// TIA Portal project "PLC_SWaT_LSTM" (V19)
// zoltan.dobrady@hotmail.com

(* hardware
DEVICE "S7-1500/ET200MP station_1"  S7-1500 station
   slot 0: "Rail_0"  Rack  6ES7 590-1***0-0AA0
   slot 1: "PLC_1"  CPU 1515F-2 PN  6ES7 515-2FM01-0AB0  V2.1
      slot 3: "CPU display_1"  6ES7591-1BA00-0AA0
      slot 32768: "PROFINET interface_1"  X1
         slot 32769: "Port_1"  X1 P1
         slot 32770: "Port_2"  X1 P2
      slot 33024: "PROFINET interface_2"  X2
         slot 33025: "Port_1"  X2 P1
*)

// ===== PLC "PLC_1"  CPU 1515F-2 PN =====

// folder: Database

DATA_BLOCK "DB_model_HS16_IW10"   // DB1
{ S7_Optimized_Access := 'TRUE' }
VERSION : 0.1
// --- Siemens Structured Format ---
   VAR
      W_i : Array[0..15, 0..39] of Real;
      W_f : Array[0..15, 0..39] of Real;
      W_g : Array[0..15, 0..39] of Real;
      W_o : Array[0..15, 0..39] of Real;
      R_i : Array[0..15, 0..15] of Real;
      R_f : Array[0..15, 0..15] of Real;
      R_g : Array[0..15, 0..15] of Real;
      R_o : Array[0..15, 0..15] of Real;
      B_i : Array[0..15] of Real;
      B_f : Array[0..15] of Real;
      B_g : Array[0..15] of Real;
      B_o : Array[0..15] of Real;
      FC_W : Array[0..39, 0..15] of Real;
      FC_B : Array[0..39] of Real;
   END_VAR
BEGIN
   W_i[0,0] := 0.03254747;
   W_i[0,1] := 0.123859;
   W_i[0,2] := 0.04015401;
   W_i[0,3] := -0.03803189;
   W_i[0,4] := 0.1759319;
   W_i[0,5] := 0.00417833;
   W_i[0,6] := -0.00157293;
   W_i[0,7] := 0.0728622;
   W_i[0,8] := 0.06175515;
   W_i[0,9] := -0.03080547;
   W_i[0,10] := 0.01361996;
   W_i[0,11] := -0.2367004;
   W_i[0,12] := 0.1251248;
   W_i[0,13] := -0.1203895;
   W_i[0,14] := 0.0523482;
   W_i[0,15] := 0.2630532;
   W_i[0,16] := -0.1147504;
   W_i[0,17] := 0.05957858;
   W_i[0,18] := -0.02271187;
   W_i[0,19] := -0.04982074;
   W_i[0,20] := 0.01270425;
   W_i[0,21] := 0.3620531;
   W_i[0,22] := -0.2914467;
   W_i[0,23] := 0.02366253;
   W_i[0,24] := -0.602429;
   W_i[0,25] := -0.5198534;
   W_i[0,26] := 0.01890776;
   W_i[0,27] := -0.4244256;
   W_i[0,28] := 0.09802054;
   W_i[0,29] := -0.2919731;
   W_i[0,30] := 0.1756448;
   W_i[0,31] := -0.06584074;
   W_i[0,32] := 0.04272554;
   W_i[0,33] := 0.06813997;
   W_i[0,34] := 0.1243908;
   W_i[0,35] := -0.2062567;
   W_i[0,36] := 0.05875245;
   W_i[0,37] := -0.2700093;
   W_i[0,38] := 0.2212317;
   W_i[0,39] := 1.454268;
   W_i[1,0] := 0.04402059;
   W_i[1,1] := 0.1007617;
   W_i[1,2] := -0.00997876;
   W_i[1,3] := 0.00796912;
   W_i[1,4] := -0.00383734;
   W_i[1,5] := -0.00800767;
   W_i[1,6] := 0.1229124;
   W_i[1,7] := 0.04417216;
   W_i[1,8] := -0.00160155;
   W_i[1,9] := -0.03973384;
   W_i[1,10] := -0.05576275;
   W_i[1,11] := 0.01415846;
   W_i[1,12] := -0.1102211;
   W_i[1,13] := 0.0361371;
   W_i[1,14] := -0.00464776;
   W_i[1,15] := -0.02071899;
   W_i[1,16] := 0.0165178;
   W_i[1,17] := -0.00011115;
   W_i[1,18] := 0.04986879;
   W_i[1,19] := -0.05042609;
   W_i[1,20] := 0.08610544;
   W_i[1,21] := 0.05673008;
   W_i[1,22] := -0.00434864;
   W_i[1,23] := 0.01197722;
   W_i[1,24] := -0.5458539;
   W_i[1,25] := -0.6899631;
   W_i[1,26] := 0.01104975;
   W_i[1,27] := 0.0182511;
   W_i[1,28] := 0.04478757;
   W_i[1,29] := -0.05586376;
   W_i[1,30] := 0.02979602;
   W_i[1,31] := 0.00707946;
   W_i[1,32] := 0.1464935;
   W_i[1,33] := 0.04832766;
   W_i[1,34] := -0.9202742;
   W_i[1,35] := -0.1918912;
   W_i[1,36] := 0.02485085;
   W_i[1,37] := -0.05241579;
   W_i[1,38] := 0.01553158;
   W_i[1,39] := -0.00394726;
   W_i[2,0] := 0.0670436;
   W_i[2,1] := -0.1175203;
   W_i[2,2] := 0.02326228;
   W_i[2,3] := -0.1431773;
   W_i[2,4] := -0.05582308;
   W_i[2,5] := 0.03605313;
   W_i[2,6] := 0.04952687;
   W_i[2,7] := -0.05419854;
   W_i[2,8] := -0.00077774;
   W_i[2,9] := 0.1769989;
   W_i[2,10] := 0.02469403;
   W_i[2,11] := 0.2849406;
   W_i[2,12] := -0.2712711;
   W_i[2,13] := -0.06837726;
   W_i[2,14] := 0.00509281;
   W_i[2,15] := 0.07467768;
   W_i[2,16] := 0.01470727;
   W_i[2,17] := 0.1139419;
   W_i[2,18] := -0.03895494;
   W_i[2,19] := 0.02999579;
   W_i[2,20] := 0.0196714;
   W_i[2,21] := 0.00220801;
   W_i[2,22] := -0.33803;
   W_i[2,23] := 0.09799825;
   W_i[2,24] := -0.5955718;
   W_i[2,25] := -0.7228485;
   W_i[2,26] := 0.07928592;
   W_i[2,27] := -0.03053538;
   W_i[2,28] := -0.1309938;
   W_i[2,29] := -0.04490006;
   W_i[2,30] := 0.05262627;
   W_i[2,31] := -0.03356259;
   W_i[2,32] := 0.06378829;
   W_i[2,33] := -0.00362085;
   W_i[2,34] := -0.6579466;
   W_i[2,35] := 0.02030313;
   W_i[2,36] := 0.05807094;
   W_i[2,37] := -0.1117615;
   W_i[2,38] := 0.09806133;
   W_i[2,39] := -0.04513157;
   W_i[3,0] := -0.03288125;
   W_i[3,1] := 0.03644303;
   W_i[3,2] := -0.02111984;
   W_i[3,3] := -0.09554495;
   W_i[3,4] := 0.471034;
   W_i[3,5] := -0.0182176;
   W_i[3,6] := -0.01296977;
   W_i[3,7] := 0.09772011;
   W_i[3,8] := 0.02375359;
   W_i[3,9] := 0.0802948;
   W_i[3,10] := 0.06341432;
   W_i[3,11] := -0.05777879;
   W_i[3,12] := 0.09200994;
   W_i[3,13] := -0.0054342;
   W_i[3,14] := -0.1107964;
   W_i[3,15] := 0.1856784;
   W_i[3,16] := -0.0179559;
   W_i[3,17] := -0.01424691;
   W_i[3,18] := 0.02418556;
   W_i[3,19] := -0.08783326;
   W_i[3,20] := 0.05560731;
   W_i[3,21] := 0.2986822;
   W_i[3,22] := -0.2220259;
   W_i[3,23] := -0.03734203;
   W_i[3,24] := 0.08825689;
   W_i[3,25] := 0.1838893;
   W_i[3,26] := 0.1152585;
   W_i[3,27] := -0.444976;
   W_i[3,28] := 0.1019801;
   W_i[3,29] := -0.4402614;
   W_i[3,30] := -0.2070405;
   W_i[3,31] := 0.00454621;
   W_i[3,32] := -0.03864358;
   W_i[3,33] := -0.1032195;
   W_i[3,34] := 0.6178231;
   W_i[3,35] := -0.01621445;
   W_i[3,36] := 0.06078746;
   W_i[3,37] := 0.07829241;
   W_i[3,38] := 0.08872399;
   W_i[3,39] := 0.01815886;
   W_i[4,0] := -0.09336383;
   W_i[4,1] := 0.00870158;
   W_i[4,2] := -0.0504511;
   W_i[4,3] := 0.0685437;
   W_i[4,4] := 0.06657482;
   W_i[4,5] := -0.04358229;
   W_i[4,6] := 0.01173393;
   W_i[4,7] := 0.02832152;
   W_i[4,8] := -0.2380867;
   W_i[4,9] := 0.2590344;
   W_i[4,10] := -0.02959821;
   W_i[4,11] := -0.1970284;
   W_i[4,12] := -0.04782372;
   W_i[4,13] := 0.00693473;
   W_i[4,14] := 0.00193878;
   W_i[4,15] := 0.03396931;
   W_i[4,16] := -0.03933699;
   W_i[4,17] := -0.09345319;
   W_i[4,18] := 0.8571873;
   W_i[4,19] := -0.208394;
   W_i[4,20] := -0.00447866;
   W_i[4,21] := -0.04350503;
   W_i[4,22] := 0.09176219;
   W_i[4,23] := 0.04992297;
   W_i[4,24] := -0.4504299;
   W_i[4,25] := 0.01641427;
   W_i[4,26] := -0.1837832;
   W_i[4,27] := 0.03955682;
   W_i[4,28] := -0.06913128;
   W_i[4,29] := 0.08025265;
   W_i[4,30] := -0.1162292;
   W_i[4,31] := 0.04558431;
   W_i[4,32] := 0.07176397;
   W_i[4,33] := -0.04032118;
   W_i[4,34] := 0.2098121;
   W_i[4,35] := -0.1125335;
   W_i[4,36] := -0.01868857;
   W_i[4,37] := -0.07242457;
   W_i[4,38] := -0.1324239;
   W_i[4,39] := -0.04244877;
   W_i[5,0] := 0.01391891;
   W_i[5,1] := -0.110183;
   W_i[5,2] := -0.00893384;
   W_i[5,3] := -0.01407803;
   W_i[5,4] := 0.08575681;
   W_i[5,5] := 0.08241521;
   W_i[5,6] := -0.06153676;
   W_i[5,7] := 0.03060099;
   W_i[5,8] := -0.03490681;
   W_i[5,9] := 0.0314279;
   W_i[5,10] := -0.02459875;
   W_i[5,11] := 0.1095907;
   W_i[5,12] := -0.02965787;
   W_i[5,13] := 0.00184801;
   W_i[5,14] := 0.02055808;
   W_i[5,15] := -0.00937524;
   W_i[5,16] := -0.01257727;
   W_i[5,17] := 0.01791891;
   W_i[5,18] := -0.0115625;
   W_i[5,19] := -0.02731706;
   W_i[5,20] := 0.08900256;
   W_i[5,21] := 0.09895428;
   W_i[5,22] := 0.02720478;
   W_i[5,23] := 0.04369688;
   W_i[5,24] := -1.906074;
   W_i[5,25] := -0.09418426;
   W_i[5,26] := -0.010597;
   W_i[5,27] := -0.09780212;
   W_i[5,28] := 0.1125583;
   W_i[5,29] := 0.08197493;
   W_i[5,30] := -0.08072126;
   W_i[5,31] := 0.03083795;
   W_i[5,32] := 0.06895962;
   W_i[5,33] := 0.00149198;
   W_i[5,34] := 0.3009818;
   W_i[5,35] := 0.1442458;
   W_i[5,36] := -0.02817895;
   W_i[5,37] := -0.08498497;
   W_i[5,38] := 0.03758771;
   W_i[5,39] := 0.01095005;
   W_i[6,0] := 0.08324189;
   W_i[6,1] := -0.2883669;
   W_i[6,2] := -0.00092833;
   W_i[6,3] := -0.00874277;
   W_i[6,4] := 0.1196982;
   W_i[6,5] := -0.1120785;
   W_i[6,6] := -0.0087709;
   W_i[6,7] := -0.03745995;
   W_i[6,8] := 0.00287988;
   W_i[6,9] := 0.00178848;
   W_i[6,10] := 0.03823818;
   W_i[6,11] := 0.02621512;
   W_i[6,12] := -0.288421;
   W_i[6,13] := -0.07084718;
   W_i[6,14] := 0.04070705;
   W_i[6,15] := -0.020424;
   W_i[6,16] := -0.00164282;
   W_i[6,17] := 0.01065832;
   W_i[6,18] := 0.00655926;
   W_i[6,19] := 0.02358968;
   W_i[6,20] := 0.1303789;
   W_i[6,21] := 0.038681;
   W_i[6,22] := -0.06235948;
   W_i[6,23] := 0.07983913;
   W_i[6,24] := -0.2428008;
   W_i[6,25] := -0.05732525;
   W_i[6,26] := 0.1651715;
   W_i[6,27] := -0.07414961;
   W_i[6,28] := 0.06032364;
   W_i[6,29] := 0.08282514;
   W_i[6,30] := -0.01358633;
   W_i[6,31] := 0.0431109;
   W_i[6,32] := 0.03472897;
   W_i[6,33] := -0.04253995;
   W_i[6,34] := 0.01447233;
   W_i[6,35] := 0.03594886;
   W_i[6,36] := -0.01385077;
   W_i[6,37] := 0.1116451;
   W_i[6,38] := 0.1253235;
   W_i[6,39] := -0.03726343;
   W_i[7,0] := 0.01927893;
   W_i[7,1] := 0.05625859;
   W_i[7,2] := 0.04672581;
   W_i[7,3] := -0.00316564;
   W_i[7,4] := 0.09401099;
   W_i[7,5] := -0.02755413;
   W_i[7,6] := -0.03952036;
   W_i[7,7] := 0.03364034;
   W_i[7,8] := 0.05500693;
   W_i[7,9] := 0.02471298;
   W_i[7,10] := 0.03820876;
   W_i[7,11] := -0.2692161;
   W_i[7,12] := -0.02231521;
   W_i[7,13] := -0.0175243;
   W_i[7,14] := 0.03934914;
   W_i[7,15] := 0.01282423;
   W_i[7,16] := -0.0871601;
   W_i[7,17] := -0.09125534;
   W_i[7,18] := 0.00613662;
   W_i[7,19] := 0.08651425;
   W_i[7,20] := -0.01288831;
   W_i[7,21] := 0.2017677;
   W_i[7,22] := -0.2016672;
   W_i[7,23] := 0.01241351;
   W_i[7,24] := -0.8755623;
   W_i[7,25] := -0.4621839;
   W_i[7,26] := 0.09773878;
   W_i[7,27] := -0.1281056;
   W_i[7,28] := 0.04194518;
   W_i[7,29] := -0.03563948;
   W_i[7,30] := 0.08049577;
   W_i[7,31] := 0.04509509;
   W_i[7,32] := -0.113328;
   W_i[7,33] := 0.1053996;
   W_i[7,34] := 0.2416716;
   W_i[7,35] := 0.04508473;
   W_i[7,36] := 0.00324964;
   W_i[7,37] := 0.2255004;
   W_i[7,38] := 0.1750992;
   W_i[7,39] := -0.7787634;
   W_i[8,0] := -0.03076644;
   W_i[8,1] := 0.03958185;
   W_i[8,2] := 0.05958826;
   W_i[8,3] := 0.00143461;
   W_i[8,4] := -0.03551066;
   W_i[8,5] := 0.0670559;
   W_i[8,6] := -0.00545013;
   W_i[8,7] := -0.1152002;
   W_i[8,8] := -0.04941865;
   W_i[8,9] := 0.00970779;
   W_i[8,10] := -0.02700928;
   W_i[8,11] := 0.1261697;
   W_i[8,12] := -0.230127;
   W_i[8,13] := -0.1321811;
   W_i[8,14] := 0.1056539;
   W_i[8,15] := 0.03265957;
   W_i[8,16] := 0.01893855;
   W_i[8,17] := 0.05783269;
   W_i[8,18] := 0.04541522;
   W_i[8,19] := -0.1756509;
   W_i[8,20] := -0.0300831;
   W_i[8,21] := 0.02609591;
   W_i[8,22] := -0.1179207;
   W_i[8,23] := -0.03097328;
   W_i[8,24] := -1.123494;
   W_i[8,25] := -0.1057856;
   W_i[8,26] := 0.1196709;
   W_i[8,27] := -0.1930985;
   W_i[8,28] := -0.04314341;
   W_i[8,29] := -0.02280886;
   W_i[8,30] := 0.09419166;
   W_i[8,31] := -0.00168002;
   W_i[8,32] := 0.170113;
   W_i[8,33] := 0.1277638;
   W_i[8,34] := 0.0079219;
   W_i[8,35] := 0.00793266;
   W_i[8,36] := 0.02933485;
   W_i[8,37] := -0.04765635;
   W_i[8,38] := -0.05385318;
   W_i[8,39] := 1.045761;
   W_i[9,0] := 0.1591891;
   W_i[9,1] := 0.04106269;
   W_i[9,2] := 0.02940365;
   W_i[9,3] := -0.02633034;
   W_i[9,4] := 0.06646424;
   W_i[9,5] := -0.06870057;
   W_i[9,6] := 0.00617184;
   W_i[9,7] := 0.01493581;
   W_i[9,8] := 0.00472299;
   W_i[9,9] := -0.1817109;
   W_i[9,10] := -0.0086358;
   W_i[9,11] := 0.1120397;
   W_i[9,12] := 0.03235663;
   W_i[9,13] := -0.00635904;
   W_i[9,14] := -0.00805719;
   W_i[9,15] := 0.03256573;
   W_i[9,16] := -0.029828;
   W_i[9,17] := 0.02432551;
   W_i[9,18] := -0.04791717;
   W_i[9,19] := -0.03479305;
   W_i[9,20] := 0.02419964;
   W_i[9,21] := -0.0080657;
   W_i[9,22] := 0.00884045;
   W_i[9,23] := 0.00822151;
   W_i[9,24] := -0.4626606;
   W_i[9,25] := -0.2415425;
   W_i[9,26] := 0.1063772;
   W_i[9,27] := 0.00555547;
   W_i[9,28] := 0.00231378;
   W_i[9,29] := 0.1730648;
   W_i[9,30] := -0.1442872;
   W_i[9,31] := -0.01611738;
   W_i[9,32] := -0.1527355;
   W_i[9,33] := -0.03995335;
   W_i[9,34] := -0.6023377;
   W_i[9,35] := -0.06071381;
   W_i[9,36] := 0.01153921;
   W_i[9,37] := 0.157252;
   W_i[9,38] := 0.04887648;
   W_i[9,39] := 0.03194974;
   W_i[10,0] := 5.71E-06;
   W_i[10,1] := 0.0292189;
   W_i[10,2] := 0.03921259;
   W_i[10,3] := -0.1034236;
   W_i[10,4] := 0.04451175;
   W_i[10,5] := -0.01788418;
   W_i[10,6] := 0.06014212;
   W_i[10,7] := -0.127616;
   W_i[10,8] := 0.1096968;
   W_i[10,9] := 0.1346427;
   W_i[10,10] := -0.07629871;
   W_i[10,11] := -1.314735;
   W_i[10,12] := 0.9704102;
   W_i[10,13] := -0.02917644;
   W_i[10,14] := 0.2685799;
   W_i[10,15] := 0.06801854;
   W_i[10,16] := -0.2241947;
   W_i[10,17] := 0.2624845;
   W_i[10,18] := -0.1694944;
   W_i[10,19] := -0.1197102;
   W_i[10,20] := -0.1591434;
   W_i[10,21] := 0.1818019;
   W_i[10,22] := -0.4487775;
   W_i[10,23] := 0.05718501;
   W_i[10,24] := 0.7740152;
   W_i[10,25] := 0.6112806;
   W_i[10,26] := 0.00735129;
   W_i[10,27] := -0.08243502;
   W_i[10,28] := -0.03729297;
   W_i[10,29] := 0.1612841;
   W_i[10,30] := -0.02351914;
   W_i[10,31] := 0.1043125;
   W_i[10,32] := 0.05746254;
   W_i[10,33] := 0.08887602;
   W_i[10,34] := -0.3910645;
   W_i[10,35] := 0.2256924;
   W_i[10,36] := -0.1320819;
   W_i[10,37] := -0.1611588;
   W_i[10,38] := 0.2708046;
   W_i[10,39] := 0.6280136;
   W_i[11,0] := -0.05849513;
   W_i[11,1] := -0.03062119;
   W_i[11,2] := -0.00411083;
   W_i[11,3] := 0.00799791;
   W_i[11,4] := 0.08333463;
   W_i[11,5] := 0.02937987;
   W_i[11,6] := 0.06844535;
   W_i[11,7] := -0.0119828;
   W_i[11,8] := 0.05660131;
   W_i[11,9] := -0.1460933;
   W_i[11,10] := -0.01666861;
   W_i[11,11] := -0.06908122;
   W_i[11,12] := 0.1548331;
   W_i[11,13] := -0.00687739;
   W_i[11,14] := 0.01971146;
   W_i[11,15] := 0.1330592;
   W_i[11,16] := -0.02189317;
   W_i[11,17] := 0.00985993;
   W_i[11,18] := -0.1488067;
   W_i[11,19] := 0.01909257;
   W_i[11,20] := 0.03714932;
   W_i[11,21] := -0.02673176;
   W_i[11,22] := -0.02788893;
   W_i[11,23] := 0.1140895;
   W_i[11,24] := -0.3711884;
   W_i[11,25] := -0.08985706;
   W_i[11,26] := -0.1102327;
   W_i[11,27] := 0.05117378;
   W_i[11,28] := 0.08547711;
   W_i[11,29] := 0.1270248;
   W_i[11,30] := 0.1054488;
   W_i[11,31] := -0.00480978;
   W_i[11,32] := 0.1614495;
   W_i[11,33] := 0.05210381;
   W_i[11,34] := -0.00085451;
   W_i[11,35] := -0.00874526;
   W_i[11,36] := -0.0616112;
   W_i[11,37] := -0.3677483;
   W_i[11,38] := 0.04212995;
   W_i[11,39] := 0.03037546;
   W_i[12,0] := 0.00629061;
   W_i[12,1] := -0.06136212;
   W_i[12,2] := -0.00718669;
   W_i[12,3] := -0.1004218;
   W_i[12,4] := 0.06293897;
   W_i[12,5] := -0.03143417;
   W_i[12,6] := -0.03538829;
   W_i[12,7] := 0.07763195;
   W_i[12,8] := -0.01023159;
   W_i[12,9] := -0.1141296;
   W_i[12,10] := -0.01354402;
   W_i[12,11] := -0.02311977;
   W_i[12,12] := 0.0279608;
   W_i[12,13] := 0.07165248;
   W_i[12,14] := -0.03632027;
   W_i[12,15] := 0.03878558;
   W_i[12,16] := -0.073125;
   W_i[12,17] := 0.01845204;
   W_i[12,18] := -0.08527449;
   W_i[12,19] := -0.00854577;
   W_i[12,20] := 0.00351815;
   W_i[12,21] := -0.1662848;
   W_i[12,22] := 0.06705266;
   W_i[12,23] := 0.1430702;
   W_i[12,24] := -0.539574;
   W_i[12,25] := -0.8721982;
   W_i[12,26] := -0.06440469;
   W_i[12,27] := 0.07379381;
   W_i[12,28] := 0.07828815;
   W_i[12,29] := 0.3882209;
   W_i[12,30] := 0.1159498;
   W_i[12,31] := 0.05581488;
   W_i[12,32] := 0.3066402;
   W_i[12,33] := 0.1275958;
   W_i[12,34] := -0.147978;
   W_i[12,35] := 0.1432935;
   W_i[12,36] := 0.2298153;
   W_i[12,37] := 0.00895516;
   W_i[12,38] := 0.2001298;
   W_i[12,39] := 0.09707437;
   W_i[13,0] := 0.07871004;
   W_i[13,1] := 0.0640982;
   W_i[13,2] := -0.00181766;
   W_i[13,3] := 0.05780525;
   W_i[13,4] := 0.2101672;
   W_i[13,5] := 0.05360549;
   W_i[13,6] := -0.0875827;
   W_i[13,7] := -0.3342811;
   W_i[13,8] := -0.09135646;
   W_i[13,9] := 0.1170631;
   W_i[13,10] := -0.0523126;
   W_i[13,11] := -0.03317479;
   W_i[13,12] := -0.403383;
   W_i[13,13] := -0.00985299;
   W_i[13,14] := 0.02202887;
   W_i[13,15] := 0.130378;
   W_i[13,16] := 0.04808246;
   W_i[13,17] := 0.04501719;
   W_i[13,18] := -0.01153503;
   W_i[13,19] := 0.03141625;
   W_i[13,20] := 0.02999944;
   W_i[13,21] := 0.01402024;
   W_i[13,22] := 0.06788336;
   W_i[13,23] := -0.09942459;
   W_i[13,24] := 0.3184399;
   W_i[13,25] := 0.1069793;
   W_i[13,26] := -0.06989229;
   W_i[13,27] := 0.1058815;
   W_i[13,28] := 0.06872193;
   W_i[13,29] := -0.1537144;
   W_i[13,30] := 0.06626805;
   W_i[13,31] := -0.0559484;
   W_i[13,32] := -0.09573574;
   W_i[13,33] := 0.05669653;
   W_i[13,34] := 0.06202357;
   W_i[13,35] := -0.1367418;
   W_i[13,36] := 0.06451428;
   W_i[13,37] := 0.1204168;
   W_i[13,38] := -0.168509;
   W_i[13,39] := 0.9775926;
   W_i[14,0] := 0.00773311;
   W_i[14,1] := -0.06673568;
   W_i[14,2] := -0.03463669;
   W_i[14,3] := -0.07830913;
   W_i[14,4] := 0.22799;
   W_i[14,5] := -0.2344869;
   W_i[14,6] := 0.1956936;
   W_i[14,7] := 0.1315334;
   W_i[14,8] := -0.1242086;
   W_i[14,9] := 0.2860397;
   W_i[14,10] := -0.09231006;
   W_i[14,11] := -0.2547791;
   W_i[14,12] := 0.1490363;
   W_i[14,13] := -0.2912802;
   W_i[14,14] := 0.1072571;
   W_i[14,15] := 0.1354038;
   W_i[14,16] := -0.09035023;
   W_i[14,17] := -0.01749873;
   W_i[14,18] := -0.4789497;
   W_i[14,19] := -0.06870104;
   W_i[14,20] := -0.1709639;
   W_i[14,21] := -0.05212005;
   W_i[14,22] := -0.1618474;
   W_i[14,23] := -0.2139406;
   W_i[14,24] := -0.7570689;
   W_i[14,25] := -0.7048593;
   W_i[14,26] := -0.3352102;
   W_i[14,27] := 0.03507431;
   W_i[14,28] := -0.1267896;
   W_i[14,29] := 0.1670964;
   W_i[14,30] := -0.0505274;
   W_i[14,31] := -0.1180039;
   W_i[14,32] := -0.0957516;
   W_i[14,33] := -0.01452094;
   W_i[14,34] := 0.00625472;
   W_i[14,35] := -0.1287756;
   W_i[14,36] := -0.06069501;
   W_i[14,37] := -0.2287704;
   W_i[14,38] := 0.1723173;
   W_i[14,39] := 1.048311;
   W_i[15,0] := 0.04376059;
   W_i[15,1] := -0.02296846;
   W_i[15,2] := 0.01713722;
   W_i[15,3] := 0.1710745;
   W_i[15,4] := 0.1736928;
   W_i[15,5] := -0.01825109;
   W_i[15,6] := -0.02258963;
   W_i[15,7] := 0.02190229;
   W_i[15,8] := -0.03702974;
   W_i[15,9] := -0.03196403;
   W_i[15,10] := 0.0826442;
   W_i[15,11] := 0.05920084;
   W_i[15,12] := -0.4280593;
   W_i[15,13] := -0.1717298;
   W_i[15,14] := 0.02115602;
   W_i[15,15] := -0.00198027;
   W_i[15,16] := 0.02912534;
   W_i[15,17] := -0.07075519;
   W_i[15,18] := -0.1174446;
   W_i[15,19] := 0.3068856;
   W_i[15,20] := 0.04301663;
   W_i[15,21] := 0.2163539;
   W_i[15,22] := -0.08966552;
   W_i[15,23] := 0.07217173;
   W_i[15,24] := -0.5324492;
   W_i[15,25] := -0.1716945;
   W_i[15,26] := -0.00556448;
   W_i[15,27] := -0.1629407;
   W_i[15,28] := 0.0326442;
   W_i[15,29] := 0.01573053;
   W_i[15,30] := -0.03329111;
   W_i[15,31] := -0.01247096;
   W_i[15,32] := 0.2100068;
   W_i[15,33] := 0.1504364;
   W_i[15,34] := -0.1697979;
   W_i[15,35] := 0.00504174;
   W_i[15,36] := 0.00267995;
   W_i[15,37] := -0.06215737;
   W_i[15,38] := 0.2148149;
   W_i[15,39] := 0.07231134;
   W_f[0,0] := -0.02091779;
   W_f[0,1] := -0.01810063;
   W_f[0,2] := 0.210087;
   W_f[0,3] := 0.09207959;
   W_f[0,4] := -0.106951;
   W_f[0,5] := -0.03611851;
   W_f[0,6] := 0.03397696;
   W_f[0,7] := 0.1654486;
   W_f[0,8] := -0.05997881;
   W_f[0,9] := -0.00453302;
   W_f[0,10] := 0.03307042;
   W_f[0,11] := 0.1420249;
   W_f[0,12] := 0.08012222;
   W_f[0,13] := -0.01528266;
   W_f[0,14] := -0.1520115;
   W_f[0,15] := -0.1571838;
   W_f[0,16] := -0.08413183;
   W_f[0,17] := 0.202225;
   W_f[0,18] := -0.01353853;
   W_f[0,19] := 0.02782044;
   W_f[0,20] := -0.04748038;
   W_f[0,21] := 0.1830429;
   W_f[0,22] := 0.312574;
   W_f[0,23] := -0.06208337;
   W_f[0,24] := 1.601337;
   W_f[0,25] := 1.519568;
   W_f[0,26] := 0.00266673;
   W_f[0,27] := 0.1218089;
   W_f[0,28] := 0.04435247;
   W_f[0,29] := 0.03200248;
   W_f[0,30] := 0.3833835;
   W_f[0,31] := 0.04435838;
   W_f[0,32] := 0.3068092;
   W_f[0,33] := 0.1323125;
   W_f[0,34] := 1.357195;
   W_f[0,35] := 0.3687007;
   W_f[0,36] := 0.08067872;
   W_f[0,37] := 0.2129946;
   W_f[0,38] := -0.02734181;
   W_f[0,39] := 0.07611577;
   W_f[1,0] := -0.388171;
   W_f[1,1] := 0.0277961;
   W_f[1,2] := -0.2651086;
   W_f[1,3] := -0.07072625;
   W_f[1,4] := 0.1196625;
   W_f[1,5] := 0.1200041;
   W_f[1,6] := -0.5084692;
   W_f[1,7] := -0.1336109;
   W_f[1,8] := -0.1377796;
   W_f[1,9] := -0.08736181;
   W_f[1,10] := 0.3113477;
   W_f[1,11] := 0.08504082;
   W_f[1,12] := 0.2114833;
   W_f[1,13] := -0.1354954;
   W_f[1,14] := -0.1227995;
   W_f[1,15] := 0.05185516;
   W_f[1,16] := -0.1474537;
   W_f[1,17] := 0.05817819;
   W_f[1,18] := 1.081658;
   W_f[1,19] := 0.1838115;
   W_f[1,20] := 0.2874206;
   W_f[1,21] := -0.2731599;
   W_f[1,22] := 0.08855448;
   W_f[1,23] := -0.09573217;
   W_f[1,24] := -0.3668332;
   W_f[1,25] := -0.6991156;
   W_f[1,26] := 0.07979747;
   W_f[1,27] := -0.1754114;
   W_f[1,28] := -0.2455159;
   W_f[1,29] := 0.1498487;
   W_f[1,30] := 0.02324941;
   W_f[1,31] := 0.07932284;
   W_f[1,32] := -0.1244244;
   W_f[1,33] := 0.02366536;
   W_f[1,34] := 0.1374529;
   W_f[1,35] := 0.4630612;
   W_f[1,36] := -0.2267325;
   W_f[1,37] := 0.07258049;
   W_f[1,38] := 0.4229668;
   W_f[1,39] := 0.1492153;
   W_f[2,0] := -0.01982149;
   W_f[2,1] := 0.03324119;
   W_f[2,2] := -0.04425151;
   W_f[2,3] := 0.08356856;
   W_f[2,4] := -0.00266197;
   W_f[2,5] := -0.01017811;
   W_f[2,6] := -0.03237398;
   W_f[2,7] := -0.00609645;
   W_f[2,8] := -0.04705935;
   W_f[2,9] := 0.03853706;
   W_f[2,10] := 0.0314042;
   W_f[2,11] := -0.1204331;
   W_f[2,12] := 0.2691576;
   W_f[2,13] := 0.04188414;
   W_f[2,14] := 0.1063143;
   W_f[2,15] := 0.05646345;
   W_f[2,16] := 0.1619761;
   W_f[2,17] := 0.2140286;
   W_f[2,18] := -0.09279267;
   W_f[2,19] := -0.0057711;
   W_f[2,20] := -0.03028176;
   W_f[2,21] := -0.05153098;
   W_f[2,22] := -0.1101711;
   W_f[2,23] := -0.01419843;
   W_f[2,24] := -0.6308476;
   W_f[2,25] := -0.4115897;
   W_f[2,26] := -0.1494104;
   W_f[2,27] := 0.04505387;
   W_f[2,28] := 0.09163468;
   W_f[2,29] := 0.2042337;
   W_f[2,30] := -0.05021087;
   W_f[2,31] := -0.05815214;
   W_f[2,32] := -0.04207016;
   W_f[2,33] := 0.2173674;
   W_f[2,34] := 0.6430734;
   W_f[2,35] := -0.1955237;
   W_f[2,36] := -0.05630085;
   W_f[2,37] := 0.0053133;
   W_f[2,38] := -0.1228282;
   W_f[2,39] := 0.5455168;
   W_f[3,0] := -0.00758014;
   W_f[3,1] := 0.00559481;
   W_f[3,2] := 0.04034248;
   W_f[3,3] := 0.02266315;
   W_f[3,4] := -0.09543922;
   W_f[3,5] := 0.03211372;
   W_f[3,6] := 0.07329436;
   W_f[3,7] := -0.04057672;
   W_f[3,8] := -0.09598581;
   W_f[3,9] := -0.00159119;
   W_f[3,10] := 0.00039486;
   W_f[3,11] := -0.00788106;
   W_f[3,12] := -0.06210583;
   W_f[3,13] := -0.01413072;
   W_f[3,14] := -0.2401386;
   W_f[3,15] := -0.07759018;
   W_f[3,16] := 0.0436046;
   W_f[3,17] := -0.2098783;
   W_f[3,18] := 0.1486036;
   W_f[3,19] := -0.02982033;
   W_f[3,20] := -0.08417022;
   W_f[3,21] := 0.08484244;
   W_f[3,22] := 0.3341856;
   W_f[3,23] := -0.01567571;
   W_f[3,24] := 1.093444;
   W_f[3,25] := 0.9772373;
   W_f[3,26] := -0.1362202;
   W_f[3,27] := -0.0995613;
   W_f[3,28] := 0.00698416;
   W_f[3,29] := 0.0005413;
   W_f[3,30] := 0.2605347;
   W_f[3,31] := -0.09947061;
   W_f[3,32] := 0.2628707;
   W_f[3,33] := 0.00611334;
   W_f[3,34] := 1.38905;
   W_f[3,35] := -0.1434975;
   W_f[3,36] := -0.00342261;
   W_f[3,37] := -0.06542191;
   W_f[3,38] := 0.1048234;
   W_f[3,39] := 0.1138595;
   W_f[4,0] := 0.2867894;
   W_f[4,1] := -0.1455002;
   W_f[4,2] := 0.2030114;
   W_f[4,3] := -0.1528496;
   W_f[4,4] := -0.1193404;
   W_f[4,5] := -0.06261637;
   W_f[4,6] := -0.09047025;
   W_f[4,7] := -0.02217131;
   W_f[4,8] := 0.3289314;
   W_f[4,9] := -0.5019218;
   W_f[4,10] := -0.02496753;
   W_f[4,11] := -0.02753776;
   W_f[4,12] := -0.3154772;
   W_f[4,13] := -0.04408565;
   W_f[4,14] := 0.05384916;
   W_f[4,15] := -0.3253689;
   W_f[4,16] := -0.01380023;
   W_f[4,17] := -0.121247;
   W_f[4,18] := 0.6214666;
   W_f[4,19] := 0.01393374;
   W_f[4,20] := 0.04359875;
   W_f[4,21] := 0.1630262;
   W_f[4,22] := -0.2102474;
   W_f[4,23] := -0.1291176;
   W_f[4,24] := -0.0868592;
   W_f[4,25] := -0.03674764;
   W_f[4,26] := 0.3087266;
   W_f[4,27] := 0.03806484;
   W_f[4,28] := 0.01020021;
   W_f[4,29] := -0.1519751;
   W_f[4,30] := 0.05839425;
   W_f[4,31] := -0.01564794;
   W_f[4,32] := -0.1834329;
   W_f[4,33] := 0.02443381;
   W_f[4,34] := 0.2140227;
   W_f[4,35] := 0.1936068;
   W_f[4,36] := 0.09160208;
   W_f[4,37] := 0.06046678;
   W_f[4,38] := -0.08968955;
   W_f[4,39] := -0.03439303;
   W_f[5,0] := -0.3995713;
   W_f[5,1] := -0.4650751;
   W_f[5,2] := -0.2646359;
   W_f[5,3] := -0.08991144;
   W_f[5,4] := -0.1660275;
   W_f[5,5] := 0.3650228;
   W_f[5,6] := -0.03514609;
   W_f[5,7] := -0.0638742;
   W_f[5,8] := 0.1263784;
   W_f[5,9] := 0.1945071;
   W_f[5,10] := -0.07852599;
   W_f[5,11] := -0.2437045;
   W_f[5,12] := -0.06879438;
   W_f[5,13] := 0.2681186;
   W_f[5,14] := 0.01808503;
   W_f[5,15] := -0.1007093;
   W_f[5,16] := 0.3104329;
   W_f[5,17] := -0.03764273;
   W_f[5,18] := -0.05466426;
   W_f[5,19] := -0.1028605;
   W_f[5,20] := -0.1891315;
   W_f[5,21] := -0.062895;
   W_f[5,22] := 0.2626143;
   W_f[5,23] := 0.1165986;
   W_f[5,24] := 2.139313;
   W_f[5,25] := 2.362694;
   W_f[5,26] := -0.4129075;
   W_f[5,27] := 0.08711372;
   W_f[5,28] := -0.06960621;
   W_f[5,29] := -0.1088286;
   W_f[5,30] := 0.02405319;
   W_f[5,31] := -0.02791615;
   W_f[5,32] := -0.03174478;
   W_f[5,33] := -0.2259803;
   W_f[5,34] := 0.02213258;
   W_f[5,35] := 0.06206211;
   W_f[5,36] := -0.220625;
   W_f[5,37] := 0.2029873;
   W_f[5,38] := 0.03730853;
   W_f[5,39] := -0.1644827;
   W_f[6,0] := 0.09157378;
   W_f[6,1] := -0.106003;
   W_f[6,2] := 0.01516851;
   W_f[6,3] := -0.09814398;
   W_f[6,4] := -0.02060772;
   W_f[6,5] := -0.1166353;
   W_f[6,6] := 0.1760547;
   W_f[6,7] := 0.1404383;
   W_f[6,8] := -0.06626645;
   W_f[6,9] := 0.0325418;
   W_f[6,10] := -0.03667779;
   W_f[6,11] := 0.03295979;
   W_f[6,12] := 0.1345612;
   W_f[6,13] := 0.1752782;
   W_f[6,14] := 0.06438499;
   W_f[6,15] := -0.1272106;
   W_f[6,16] := -0.2878087;
   W_f[6,17] := 0.1161476;
   W_f[6,18] := -0.2311435;
   W_f[6,19] := -0.07521003;
   W_f[6,20] := -0.1416016;
   W_f[6,21] := 0.1268703;
   W_f[6,22] := 0.3855781;
   W_f[6,23] := -0.1290094;
   W_f[6,24] := 1.145507;
   W_f[6,25] := 1.206513;
   W_f[6,26] := 0.01718643;
   W_f[6,27] := -0.2014013;
   W_f[6,28] := -0.03907681;
   W_f[6,29] := -1.031836;
   W_f[6,30] := 0.1329869;
   W_f[6,31] := -0.05304611;
   W_f[6,32] := 0.2754238;
   W_f[6,33] := 0.484001;
   W_f[6,34] := 0.8730348;
   W_f[6,35] := -0.2791631;
   W_f[6,36] := 0.09285419;
   W_f[6,37] := -0.00086587;
   W_f[6,38] := 0.2140355;
   W_f[6,39] := 0.01036415;
   W_f[7,0] := -0.00185265;
   W_f[7,1] := 0.07858364;
   W_f[7,2] := 0.00610039;
   W_f[7,3] := 0.06575946;
   W_f[7,4] := -0.0810083;
   W_f[7,5] := 0.00321988;
   W_f[7,6] := 0.07597861;
   W_f[7,7] := -0.1263862;
   W_f[7,8] := 0.1467239;
   W_f[7,9] := 0.04145058;
   W_f[7,10] := 0.03552409;
   W_f[7,11] := -0.4200411;
   W_f[7,12] := 0.2535799;
   W_f[7,13] := -0.08330481;
   W_f[7,14] := -0.08974353;
   W_f[7,15] := -0.1051762;
   W_f[7,16] := -0.3822444;
   W_f[7,17] := -0.4579986;
   W_f[7,18] := -0.06309059;
   W_f[7,19] := -0.3079986;
   W_f[7,20] := -0.08522949;
   W_f[7,21] := -0.06581733;
   W_f[7,22] := 0.2580513;
   W_f[7,23] := 0.02311642;
   W_f[7,24] := 0.9095069;
   W_f[7,25] := 1.188896;
   W_f[7,26] := -0.1154661;
   W_f[7,27] := -0.1087225;
   W_f[7,28] := -0.08876549;
   W_f[7,29] := 0.00109644;
   W_f[7,30] := 0.2337219;
   W_f[7,31] := -0.1376933;
   W_f[7,32] := 0.1659716;
   W_f[7,33] := 0.04170239;
   W_f[7,34] := 1.311337;
   W_f[7,35] := -0.1188877;
   W_f[7,36] := 0.04907094;
   W_f[7,37] := 0.1402612;
   W_f[7,38] := 0.1255982;
   W_f[7,39] := -1.274189;
   W_f[8,0] := 0.12556;
   W_f[8,1] := -0.1031576;
   W_f[8,2] := 0.03551091;
   W_f[8,3] := -0.03898631;
   W_f[8,4] := -0.1320676;
   W_f[8,5] := 0.07454634;
   W_f[8,6] := 0.1020655;
   W_f[8,7] := 0.01262685;
   W_f[8,8] := -0.00534601;
   W_f[8,9] := -0.00536494;
   W_f[8,10] := -0.04092396;
   W_f[8,11] := -0.3869237;
   W_f[8,12] := 0.03422466;
   W_f[8,13] := 0.02580789;
   W_f[8,14] := 0.2689887;
   W_f[8,15] := -0.2494489;
   W_f[8,16] := -0.02722716;
   W_f[8,17] := -0.1010804;
   W_f[8,18] := 0.5424435;
   W_f[8,19] := -0.2312066;
   W_f[8,20] := -0.04103015;
   W_f[8,21] := -0.1674081;
   W_f[8,22] := 0.1389381;
   W_f[8,23] := -0.04656294;
   W_f[8,24] := 0.531742;
   W_f[8,25] := 0.7430941;
   W_f[8,26] := -0.00084738;
   W_f[8,27] := -0.04600925;
   W_f[8,28] := -0.1588;
   W_f[8,29] := 0.08535929;
   W_f[8,30] := 0.1022129;
   W_f[8,31] := -0.03335671;
   W_f[8,32] := 0.03138823;
   W_f[8,33] := -0.02403146;
   W_f[8,34] := 0.8330596;
   W_f[8,35] := -0.07033388;
   W_f[8,36] := -0.1749986;
   W_f[8,37] := 0.0922937;
   W_f[8,38] := -0.1766868;
   W_f[8,39] := 0.141985;
   W_f[9,0] := -0.08198071;
   W_f[9,1] := 0.03835172;
   W_f[9,2] := 1.020265;
   W_f[9,3] := -0.1529395;
   W_f[9,4] := -0.1617989;
   W_f[9,5] := 0.03072036;
   W_f[9,6] := -0.09759208;
   W_f[9,7] := -0.07946933;
   W_f[9,8] := -0.6549187;
   W_f[9,9] := 0.2455487;
   W_f[9,10] := -0.00084776;
   W_f[9,11] := -0.02393647;
   W_f[9,12] := -0.1103576;
   W_f[9,13] := 0.05757844;
   W_f[9,14] := 0.00252463;
   W_f[9,15] := -0.04278835;
   W_f[9,16] := -0.01363701;
   W_f[9,17] := 0.03181182;
   W_f[9,18] := 0.2954217;
   W_f[9,19] := 0.1868071;
   W_f[9,20] := -0.1459624;
   W_f[9,21] := 0.04626612;
   W_f[9,22] := -0.4959656;
   W_f[9,23] := -0.298828;
   W_f[9,24] := -0.05025842;
   W_f[9,25] := -0.2492222;
   W_f[9,26] := 0.2277043;
   W_f[9,27] := -0.077122;
   W_f[9,28] := -0.1601862;
   W_f[9,29] := -0.360285;
   W_f[9,30] := -0.1589459;
   W_f[9,31] := 0.07634185;
   W_f[9,32] := -0.1424809;
   W_f[9,33] := 0.4724371;
   W_f[9,34] := 0.3722708;
   W_f[9,35] := 0.08862774;
   W_f[9,36] := 0.1802045;
   W_f[9,37] := -0.4637271;
   W_f[9,38] := 0.1014335;
   W_f[9,39] := 0.0325746;
   W_f[10,0] := 0.01476683;
   W_f[10,1] := 0.0891594;
   W_f[10,2] := 0.09493639;
   W_f[10,3] := 0.0092164;
   W_f[10,4] := -0.4010172;
   W_f[10,5] := -0.09464957;
   W_f[10,6] := -0.04691195;
   W_f[10,7] := -0.02866868;
   W_f[10,8] := -0.04315028;
   W_f[10,9] := -0.1709383;
   W_f[10,10] := -0.00073274;
   W_f[10,11] := -0.2750555;
   W_f[10,12] := 0.3360567;
   W_f[10,13] := -0.2203442;
   W_f[10,14] := 0.2416514;
   W_f[10,15] := -0.2352184;
   W_f[10,16] := -0.00154005;
   W_f[10,17] := -0.00158511;
   W_f[10,18] := 0.1191233;
   W_f[10,19] := -0.02448388;
   W_f[10,20] := -0.2385904;
   W_f[10,21] := -0.05945824;
   W_f[10,22] := 0.01714438;
   W_f[10,23] := -0.1828551;
   W_f[10,24] := 1.57859;
   W_f[10,25] := 1.894226;
   W_f[10,26] := 0.09559432;
   W_f[10,27] := -0.273827;
   W_f[10,28] := -0.2814649;
   W_f[10,29] := 0.04344108;
   W_f[10,30] := 0.08430442;
   W_f[10,31] := 0.1357144;
   W_f[10,32] := 0.03089454;
   W_f[10,33] := 0.1987186;
   W_f[10,34] := 0.1212473;
   W_f[10,35] := 0.1387797;
   W_f[10,36] := 0.2638152;
   W_f[10,37] := 0.00209056;
   W_f[10,38] := -0.08942132;
   W_f[10,39] := -0.4494387;
   W_f[11,0] := 0.04211291;
   W_f[11,1] := -0.02505053;
   W_f[11,2] := 0.08745301;
   W_f[11,3] := -0.04265523;
   W_f[11,4] := -0.2127612;
   W_f[11,5] := 0.01322894;
   W_f[11,6] := 0.1062051;
   W_f[11,7] := 0.01512342;
   W_f[11,8] := -0.07057641;
   W_f[11,9] := 0.1239847;
   W_f[11,10] := -0.1409187;
   W_f[11,11] := -0.0726796;
   W_f[11,12] := 0.00417219;
   W_f[11,13] := -0.01783882;
   W_f[11,14] := 0.01799064;
   W_f[11,15] := -0.05493079;
   W_f[11,16] := -0.05114271;
   W_f[11,17] := -0.03128599;
   W_f[11,18] := 0.03801877;
   W_f[11,19] := -0.01814952;
   W_f[11,20] := -0.09758195;
   W_f[11,21] := -0.04573784;
   W_f[11,22] := -0.03167154;
   W_f[11,23] := -0.08901857;
   W_f[11,24] := -0.2217392;
   W_f[11,25] := 0.3994405;
   W_f[11,26] := 0.0512911;
   W_f[11,27] := 0.05733421;
   W_f[11,28] := -0.1220476;
   W_f[11,29] := 0.2530152;
   W_f[11,30] := -0.01943143;
   W_f[11,31] := 0.06523979;
   W_f[11,32] := -0.1965705;
   W_f[11,33] := 0.010429;
   W_f[11,34] := 0.1933591;
   W_f[11,35] := -0.02032585;
   W_f[11,36] := -0.05446678;
   W_f[11,37] := 0.1093058;
   W_f[11,38] := -0.05791799;
   W_f[11,39] := 0.3272165;
   W_f[12,0] := 0.0583974;
   W_f[12,1] := 0.06337267;
   W_f[12,2] := 0.05269343;
   W_f[12,3] := -0.02425898;
   W_f[12,4] := 0.0733385;
   W_f[12,5] := 0.01520942;
   W_f[12,6] := 0.03044897;
   W_f[12,7] := 0.1151135;
   W_f[12,8] := 0.03681342;
   W_f[12,9] := -0.0168035;
   W_f[12,10] := 0.04408923;
   W_f[12,11] := 0.08383411;
   W_f[12,12] := -0.01220268;
   W_f[12,13] := 0.0539641;
   W_f[12,14] := -0.07032214;
   W_f[12,15] := -0.00997462;
   W_f[12,16] := -0.06021495;
   W_f[12,17] := -0.01422043;
   W_f[12,18] := -0.00584967;
   W_f[12,19] := 0.05498984;
   W_f[12,20] := -0.0921667;
   W_f[12,21] := 0.1078821;
   W_f[12,22] := 0.09067565;
   W_f[12,23] := -0.09486815;
   W_f[12,24] := -0.8760142;
   W_f[12,25] := 0.543728;
   W_f[12,26] := 0.0473772;
   W_f[12,27] := -0.1004083;
   W_f[12,28] := 0.07258554;
   W_f[12,29] := 0.07306878;
   W_f[12,30] := -0.1469819;
   W_f[12,31] := 0.01059632;
   W_f[12,32] := 0.01764544;
   W_f[12,33] := -0.04630747;
   W_f[12,34] := 0.04829778;
   W_f[12,35] := -0.00637231;
   W_f[12,36] := 0.3430251;
   W_f[12,37] := 0.1221798;
   W_f[12,38] := 0.04078831;
   W_f[12,39] := 0.02011232;
   W_f[13,0] := 0.1598776;
   W_f[13,1] := 0.08477814;
   W_f[13,2] := -0.1199006;
   W_f[13,3] := -0.2151837;
   W_f[13,4] := 0.04422749;
   W_f[13,5] := 0.1643971;
   W_f[13,6] := -0.01991516;
   W_f[13,7] := 0.01602156;
   W_f[13,8] := -0.134406;
   W_f[13,9] := 0.0432152;
   W_f[13,10] := 0.1258369;
   W_f[13,11] := 0.03486055;
   W_f[13,12] := 0.1840334;
   W_f[13,13] := 0.05531228;
   W_f[13,14] := -0.05205994;
   W_f[13,15] := -0.1417992;
   W_f[13,16] := 0.2145569;
   W_f[13,17] := -0.03670088;
   W_f[13,18] := 0.05554622;
   W_f[13,19] := -0.0701214;
   W_f[13,20] := 0.05645064;
   W_f[13,21] := 0.04904451;
   W_f[13,22] := 0.1227407;
   W_f[13,23] := -0.1391225;
   W_f[13,24] := 1.281417;
   W_f[13,25] := 1.152952;
   W_f[13,26] := 0.02036783;
   W_f[13,27] := 6.46E-06;
   W_f[13,28] := 0.05594068;
   W_f[13,29] := 0.1138421;
   W_f[13,30] := 0.2391586;
   W_f[13,31] := 0.04423625;
   W_f[13,32] := 0.3790507;
   W_f[13,33] := 0.01350218;
   W_f[13,34] := 0.907777;
   W_f[13,35] := -0.01705103;
   W_f[13,36] := 0.08728553;
   W_f[13,37] := 0.1376872;
   W_f[13,38] := 0.05409899;
   W_f[13,39] := 0.5876323;
   W_f[14,0] := -0.1830878;
   W_f[14,1] := 0.00258858;
   W_f[14,2] := -0.05409549;
   W_f[14,3] := 0.4265317;
   W_f[14,4] := -0.1661472;
   W_f[14,5] := -0.06032855;
   W_f[14,6] := 0.09126755;
   W_f[14,7] := -0.1622344;
   W_f[14,8] := -0.0415544;
   W_f[14,9] := -0.03031821;
   W_f[14,10] := -0.07388397;
   W_f[14,11] := -0.1665972;
   W_f[14,12] := 0.1223991;
   W_f[14,13] := -0.1334893;
   W_f[14,14] := -0.06961614;
   W_f[14,15] := -0.04957403;
   W_f[14,16] := 0.0298849;
   W_f[14,17] := -0.1339389;
   W_f[14,18] := -0.04285705;
   W_f[14,19] := -0.08629614;
   W_f[14,20] := -0.1532967;
   W_f[14,21] := 0.04812383;
   W_f[14,22] := -0.03088393;
   W_f[14,23] := -0.04624541;
   W_f[14,24] := -0.07781153;
   W_f[14,25] := -0.8319644;
   W_f[14,26] := 0.1015401;
   W_f[14,27] := 0.04807844;
   W_f[14,28] := 0.08697836;
   W_f[14,29] := -0.3099394;
   W_f[14,30] := 0.02526759;
   W_f[14,31] := 0.06875665;
   W_f[14,32] := 0.05270454;
   W_f[14,33] := 0.08052166;
   W_f[14,34] := 0.07316659;
   W_f[14,35] := -0.2259305;
   W_f[14,36] := -0.0360414;
   W_f[14,37] := -0.1107528;
   W_f[14,38] := 0.1422287;
   W_f[14,39] := 0.1191253;
   W_f[15,0] := 0.06860624;
   W_f[15,1] := 0.2116713;
   W_f[15,2] := -0.1070077;
   W_f[15,3] := -0.1796377;
   W_f[15,4] := 0.06190439;
   W_f[15,5] := 0.1118638;
   W_f[15,6] := 0.2123804;
   W_f[15,7] := 0.04805397;
   W_f[15,8] := 0.02383129;
   W_f[15,9] := -0.08112741;
   W_f[15,10] := -0.00035556;
   W_f[15,11] := -0.00759834;
   W_f[15,12] := 0.04278949;
   W_f[15,13] := -0.01575772;
   W_f[15,14] := -0.06780741;
   W_f[15,15] := 0.07988951;
   W_f[15,16] := 0.3583542;
   W_f[15,17] := -0.1143483;
   W_f[15,18] := 0.06204842;
   W_f[15,19] := -0.1630864;
   W_f[15,20] := -0.08014372;
   W_f[15,21] := 0.09970582;
   W_f[15,22] := -0.01455338;
   W_f[15,23] := -0.09048357;
   W_f[15,24] := 1.480857;
   W_f[15,25] := 1.437098;
   W_f[15,26] := -0.04126001;
   W_f[15,27] := 0.03295555;
   W_f[15,28] := -0.0889762;
   W_f[15,29] := 0.1496947;
   W_f[15,30] := 0.1286354;
   W_f[15,31] := -0.01891266;
   W_f[15,32] := -0.08377147;
   W_f[15,33] := 0.04984247;
   W_f[15,34] := 0.7321002;
   W_f[15,35] := -0.07470711;
   W_f[15,36] := 0.01260767;
   W_f[15,37] := -0.02138078;
   W_f[15,38] := 0.01280809;
   W_f[15,39] := 0.1211099;
   W_g[0,0] := 0.1320454;
   W_g[0,1] := -0.07179091;
   W_g[0,2] := 0.1304129;
   W_g[0,3] := -0.01710966;
   W_g[0,4] := 0.08717188;
   W_g[0,5] := -0.03005558;
   W_g[0,6] := 0.02608494;
   W_g[0,7] := -0.02178418;
   W_g[0,8] := -0.02002059;
   W_g[0,9] := -0.01907159;
   W_g[0,10] := -0.07584066;
   W_g[0,11] := -0.0276128;
   W_g[0,12] := -0.03857584;
   W_g[0,13] := -0.01737243;
   W_g[0,14] := -0.1033841;
   W_g[0,15] := -0.00566125;
   W_g[0,16] := -0.01846444;
   W_g[0,17] := -0.09568264;
   W_g[0,18] := 0.01344434;
   W_g[0,19] := -0.04545733;
   W_g[0,20] := -0.07012872;
   W_g[0,21] := -0.2265758;
   W_g[0,22] := -0.0013438;
   W_g[0,23] := 0.0140279;
   W_g[0,24] := 0.05787951;
   W_g[0,25] := 0.3332284;
   W_g[0,26] := 0.1338745;
   W_g[0,27] := -0.284954;
   W_g[0,28] := 0.08640742;
   W_g[0,29] := 0.00553245;
   W_g[0,30] := 0.00379307;
   W_g[0,31] := 0.00939364;
   W_g[0,32] := -0.0225928;
   W_g[0,33] := -0.03415785;
   W_g[0,34] := 0.4156659;
   W_g[0,35] := -0.02096383;
   W_g[0,36] := -0.0417503;
   W_g[0,37] := -0.04161927;
   W_g[0,38] := 0.04176929;
   W_g[0,39] := -0.02666814;
   W_g[1,0] := 0.1003403;
   W_g[1,1] := 0.02818905;
   W_g[1,2] := 0.08966444;
   W_g[1,3] := 0.02384869;
   W_g[1,4] := -0.00957148;
   W_g[1,5] := 0.0225874;
   W_g[1,6] := 0.2189841;
   W_g[1,7] := 0.03297459;
   W_g[1,8] := 0.02741309;
   W_g[1,9] := 0.03524271;
   W_g[1,10] := -0.09459055;
   W_g[1,11] := 0.00226336;
   W_g[1,12] := -0.03214818;
   W_g[1,13] := 0.09925831;
   W_g[1,14] := 0.03271784;
   W_g[1,15] := -0.00993501;
   W_g[1,16] := 0.04625125;
   W_g[1,17] := -0.01382133;
   W_g[1,18] := 0.141697;
   W_g[1,19] := -0.06103647;
   W_g[1,20] := -0.2125344;
   W_g[1,21] := 0.1183949;
   W_g[1,22] := -0.01691977;
   W_g[1,23] := 0.05358729;
   W_g[1,24] := -0.3285331;
   W_g[1,25] := -0.4942485;
   W_g[1,26] := -0.08112237;
   W_g[1,27] := 0.1249737;
   W_g[1,28] := 0.1749274;
   W_g[1,29] := 0.05923015;
   W_g[1,30] := -0.03070631;
   W_g[1,31] := -0.0160953;
   W_g[1,32] := 0.0128262;
   W_g[1,33] := 0.00597268;
   W_g[1,34] := -0.4454135;
   W_g[1,35] := 0.04373179;
   W_g[1,36] := 0.07117015;
   W_g[1,37] := -0.05477969;
   W_g[1,38] := -0.1148913;
   W_g[1,39] := -0.05603904;
   W_g[2,0] := -0.03656583;
   W_g[2,1] := 0.08601304;
   W_g[2,2] := -0.02144271;
   W_g[2,3] := -0.00415884;
   W_g[2,4] := 0.05374509;
   W_g[2,5] := 0.01513857;
   W_g[2,6] := 0.00031003;
   W_g[2,7] := -0.00429267;
   W_g[2,8] := 0.0024794;
   W_g[2,9] := -0.02802207;
   W_g[2,10] := 0.00567887;
   W_g[2,11] := 0.07285577;
   W_g[2,12] := 0.06949551;
   W_g[2,13] := -0.06609099;
   W_g[2,14] := 0.02675425;
   W_g[2,15] := 0.05979875;
   W_g[2,16] := 0.1882337;
   W_g[2,17] := 0.1013563;
   W_g[2,18] := -0.01730143;
   W_g[2,19] := 0.07176489;
   W_g[2,20] := -0.00487325;
   W_g[2,21] := -0.01244247;
   W_g[2,22] := 0.07138075;
   W_g[2,23] := -0.08855219;
   W_g[2,24] := 0.6691746;
   W_g[2,25] := 0.4066471;
   W_g[2,26] := 0.05317146;
   W_g[2,27] := -0.03753066;
   W_g[2,28] := 0.04217075;
   W_g[2,29] := -0.08696262;
   W_g[2,30] := 0.0727913;
   W_g[2,31] := 0.04612178;
   W_g[2,32] := 0.06409022;
   W_g[2,33] := 0.01605693;
   W_g[2,34] := 0.1564854;
   W_g[2,35] := 0.1177737;
   W_g[2,36] := -0.03577918;
   W_g[2,37] := -0.02626175;
   W_g[2,38] := -0.2925088;
   W_g[2,39] := -0.1730511;
   W_g[3,0] := 0.0353583;
   W_g[3,1] := -0.1049412;
   W_g[3,2] := 0.03618518;
   W_g[3,3] := -0.03134191;
   W_g[3,4] := -0.2461421;
   W_g[3,5] := 0.1266218;
   W_g[3,6] := 0.06337537;
   W_g[3,7] := -0.035273;
   W_g[3,8] := -0.03651504;
   W_g[3,9] := -0.03074392;
   W_g[3,10] := -0.05727396;
   W_g[3,11] := -0.02935094;
   W_g[3,12] := -0.03621458;
   W_g[3,13] := -0.01833671;
   W_g[3,14] := -0.1685012;
   W_g[3,15] := -0.00882464;
   W_g[3,16] := -0.02389451;
   W_g[3,17] := -0.07828564;
   W_g[3,18] := 0.02588245;
   W_g[3,19] := -0.04996347;
   W_g[3,20] := -0.03450434;
   W_g[3,21] := 0.08713186;
   W_g[3,22] := 0.04250673;
   W_g[3,23] := 0.0231547;
   W_g[3,24] := 0.2406025;
   W_g[3,25] := -0.04010823;
   W_g[3,26] := -0.04215078;
   W_g[3,27] := 0.0426458;
   W_g[3,28] := -0.2496434;
   W_g[3,29] := -0.019585;
   W_g[3,30] := 0.03981116;
   W_g[3,31] := 0.05331163;
   W_g[3,32] := 0.02955173;
   W_g[3,33] := 0.03688915;
   W_g[3,34] := -0.07779746;
   W_g[3,35] := 0.04131736;
   W_g[3,36] := -0.09415401;
   W_g[3,37] := 0.02781735;
   W_g[3,38] := -0.01530841;
   W_g[3,39] := -0.103936;
   W_g[4,0] := 0.07740436;
   W_g[4,1] := -0.07530216;
   W_g[4,2] := 0.08100316;
   W_g[4,3] := -0.03866265;
   W_g[4,4] := -0.124116;
   W_g[4,5] := -0.06374057;
   W_g[4,6] := -0.06540763;
   W_g[4,7] := -0.05087971;
   W_g[4,8] := -0.02486523;
   W_g[4,9] := -0.00432705;
   W_g[4,10] := -0.02001161;
   W_g[4,11] := -0.2260205;
   W_g[4,12] := -0.2710404;
   W_g[4,13] := -0.04622217;
   W_g[4,14] := 0.03693646;
   W_g[4,15] := -0.2228938;
   W_g[4,16] := -0.03339233;
   W_g[4,17] := -0.1039548;
   W_g[4,18] := -0.6776975;
   W_g[4,19] := -0.1070111;
   W_g[4,20] := -0.00507321;
   W_g[4,21] := 0.06153874;
   W_g[4,22] := -0.05829039;
   W_g[4,23] := -0.03399877;
   W_g[4,24] := 0.02580869;
   W_g[4,25] := -0.05605169;
   W_g[4,26] := 0.02870816;
   W_g[4,27] := 0.09912029;
   W_g[4,28] := -0.08475526;
   W_g[4,29] := 0.02515182;
   W_g[4,30] := -0.06613169;
   W_g[4,31] := -0.01619294;
   W_g[4,32] := -0.07978069;
   W_g[4,33] := -0.02161121;
   W_g[4,34] := -0.01309834;
   W_g[4,35] := -0.0583593;
   W_g[4,36] := 0.02740471;
   W_g[4,37] := -0.06427267;
   W_g[4,38] := -0.1435904;
   W_g[4,39] := -0.04779189;
   W_g[5,0] := 0.07845761;
   W_g[5,1] := 0.122912;
   W_g[5,2] := 0.09020026;
   W_g[5,3] := -0.05951332;
   W_g[5,4] := -0.1863579;
   W_g[5,5] := -0.6706011;
   W_g[5,6] := -0.09371807;
   W_g[5,7] := -0.0624865;
   W_g[5,8] := -0.05328716;
   W_g[5,9] := -0.05699488;
   W_g[5,10] := -0.2100334;
   W_g[5,11] := -0.04094445;
   W_g[5,12] := -0.03951516;
   W_g[5,13] := 0.01896183;
   W_g[5,14] := 0.05772699;
   W_g[5,15] := -0.03484442;
   W_g[5,16] := -0.08915464;
   W_g[5,17] := -0.03359089;
   W_g[5,18] := 0.05330428;
   W_g[5,19] := -0.04913564;
   W_g[5,20] := -0.02437795;
   W_g[5,21] := -0.03660732;
   W_g[5,22] := 0.05388405;
   W_g[5,23] := 0.03580718;
   W_g[5,24] := 0.6679524;
   W_g[5,25] := 0.3846368;
   W_g[5,26] := 0.03221167;
   W_g[5,27] := -0.09449711;
   W_g[5,28] := -0.2133287;
   W_g[5,29] := -0.1070377;
   W_g[5,30] := 0.0486634;
   W_g[5,31] := 0.04555348;
   W_g[5,32] := 0.03119684;
   W_g[5,33] := 0.02472051;
   W_g[5,34] := -0.00109696;
   W_g[5,35] := 0.00976827;
   W_g[5,36] := -0.04086661;
   W_g[5,37] := 0.01402589;
   W_g[5,38] := 0.01088466;
   W_g[5,39] := 0.05395384;
   W_g[6,0] := -0.09459254;
   W_g[6,1] := -0.3465888;
   W_g[6,2] := -0.1204124;
   W_g[6,3] := 0.1131463;
   W_g[6,4] := 0.07203985;
   W_g[6,5] := -0.09553758;
   W_g[6,6] := -0.03457065;
   W_g[6,7] := 0.1258941;
   W_g[6,8] := 0.09656766;
   W_g[6,9] := 0.1205588;
   W_g[6,10] := 0.01646312;
   W_g[6,11] := -0.06715041;
   W_g[6,12] := -0.08268934;
   W_g[6,13] := -0.01733059;
   W_g[6,14] := 0.05910295;
   W_g[6,15] := -0.07129493;
   W_g[6,16] := -0.06239159;
   W_g[6,17] := -0.06886618;
   W_g[6,18] := 0.04810062;
   W_g[6,19] := -0.0965384;
   W_g[6,20] := 0.1695917;
   W_g[6,21] := -0.00798076;
   W_g[6,22] := 0.00821575;
   W_g[6,23] := 0.1049357;
   W_g[6,24] := 0.06085224;
   W_g[6,25] := 0.05369381;
   W_g[6,26] := -0.0201011;
   W_g[6,27] := 0.00523888;
   W_g[6,28] := -0.05049808;
   W_g[6,29] := 0.04111513;
   W_g[6,30] := 0.01227053;
   W_g[6,31] := 0.0204126;
   W_g[6,32] := -0.00532885;
   W_g[6,33] := -0.00633689;
   W_g[6,34] := -0.01163891;
   W_g[6,35] := 0.0326525;
   W_g[6,36] := -0.08721739;
   W_g[6,37] := 0.02508505;
   W_g[6,38] := -0.1394214;
   W_g[6,39] := -0.03058173;
   W_g[7,0] := 0.1329033;
   W_g[7,1] := -0.2278838;
   W_g[7,2] := 0.1442183;
   W_g[7,3] := -0.04011448;
   W_g[7,4] := -0.0098335;
   W_g[7,5] := 0.06002469;
   W_g[7,6] := 0.01148172;
   W_g[7,7] := -0.03318439;
   W_g[7,8] := -0.04474748;
   W_g[7,9] := -0.03664961;
   W_g[7,10] := -0.05171043;
   W_g[7,11] := 0.1588942;
   W_g[7,12] := 0.1881699;
   W_g[7,13] := 0.03320323;
   W_g[7,14] := 0.08849441;
   W_g[7,15] := 0.1089842;
   W_g[7,16] := -0.1042355;
   W_g[7,17] := 0.2178806;
   W_g[7,18] := -0.09352972;
   W_g[7,19] := 0.2286143;
   W_g[7,20] := 0.01804306;
   W_g[7,21] := 0.02883035;
   W_g[7,22] := 0.02334912;
   W_g[7,23] := 0.0097255;
   W_g[7,24] := 0.09000973;
   W_g[7,25] := 0.2379663;
   W_g[7,26] := -0.00529223;
   W_g[7,27] := 0.02389492;
   W_g[7,28] := 0.01771568;
   W_g[7,29] := 0.03995743;
   W_g[7,30] := 0.0237428;
   W_g[7,31] := 0.00652028;
   W_g[7,32] := 0.0237922;
   W_g[7,33] := 0.01227521;
   W_g[7,34] := -0.02105843;
   W_g[7,35] := 0.02154919;
   W_g[7,36] := -0.01575272;
   W_g[7,37] := -0.01810107;
   W_g[7,38] := -0.00772995;
   W_g[7,39] := -0.2820103;
   W_g[8,0] := 0.01713815;
   W_g[8,1] := -0.00229361;
   W_g[8,2] := 0.01726119;
   W_g[8,3] := -0.02061658;
   W_g[8,4] := -0.04641379;
   W_g[8,5] := 0.04689364;
   W_g[8,6] := 0.00514349;
   W_g[8,7] := -0.02527735;
   W_g[8,8] := -0.02019661;
   W_g[8,9] := -0.01965989;
   W_g[8,10] := -0.02106753;
   W_g[8,11] := -0.1810846;
   W_g[8,12] := -0.1747753;
   W_g[8,13] := -0.07262667;
   W_g[8,14] := 0.09604074;
   W_g[8,15] := -0.2233989;
   W_g[8,16] := -0.01457437;
   W_g[8,17] := 0.1895211;
   W_g[8,18] := 0.09061687;
   W_g[8,19] := -0.1659747;
   W_g[8,20] := -0.02462232;
   W_g[8,21] := -0.0811555;
   W_g[8,22] := 0.02058986;
   W_g[8,23] := -0.05404805;
   W_g[8,24] := -0.07197467;
   W_g[8,25] := -0.2429945;
   W_g[8,26] := 0.03455175;
   W_g[8,27] := -0.1281454;
   W_g[8,28] := -0.1244678;
   W_g[8,29] := -0.0707626;
   W_g[8,30] := 0.03440274;
   W_g[8,31] := 0.02760479;
   W_g[8,32] := -0.00320816;
   W_g[8,33] := -0.00195394;
   W_g[8,34] := -0.06706773;
   W_g[8,35] := -0.03631235;
   W_g[8,36] := -0.0461507;
   W_g[8,37] := 0.02211455;
   W_g[8,38] := 0.00710197;
   W_g[8,39] := 0.06994114;
   W_g[9,0] := -0.2685941;
   W_g[9,1] := -0.1633901;
   W_g[9,2] := -0.3089246;
   W_g[9,3] := -0.1282196;
   W_g[9,4] := 0.01028809;
   W_g[9,5] := -0.05689346;
   W_g[9,6] := 0.131765;
   W_g[9,7] := -0.1136668;
   W_g[9,8] := -0.1350522;
   W_g[9,9] := -0.1341046;
   W_g[9,10] := -0.2973659;
   W_g[9,11] := 0.03893382;
   W_g[9,12] := 0.03934914;
   W_g[9,13] := 0.01418684;
   W_g[9,14] := 0.01693503;
   W_g[9,15] := 0.04444136;
   W_g[9,16] := 0.07951424;
   W_g[9,17] := 0.00626671;
   W_g[9,18] := -0.06104251;
   W_g[9,19] := 0.04594292;
   W_g[9,20] := -0.02836513;
   W_g[9,21] := 0.0397499;
   W_g[9,22] := -0.02700124;
   W_g[9,23] := 0.02002714;
   W_g[9,24] := -0.5077276;
   W_g[9,25] := -0.2546269;
   W_g[9,26] := -0.03511217;
   W_g[9,27] := 0.04529352;
   W_g[9,28] := 0.04820129;
   W_g[9,29] := 0.09988645;
   W_g[9,30] := -0.01425081;
   W_g[9,31] := -0.01030078;
   W_g[9,32] := -0.01629252;
   W_g[9,33] := -0.00994037;
   W_g[9,34] := -0.5942311;
   W_g[9,35] := 0.03158842;
   W_g[9,36] := -0.08265782;
   W_g[9,37] := -0.0352644;
   W_g[9,38] := -0.00322891;
   W_g[9,39] := -0.00800959;
   W_g[10,0] := -0.03213325;
   W_g[10,1] := -0.00863164;
   W_g[10,2] := -0.03062097;
   W_g[10,3] := 0.0125538;
   W_g[10,4] := 0.1017359;
   W_g[10,5] := -0.04505892;
   W_g[10,6] := -0.00103756;
   W_g[10,7] := 0.01735601;
   W_g[10,8] := 0.01301922;
   W_g[10,9] := 0.0136564;
   W_g[10,10] := 0.00548952;
   W_g[10,11] := -0.00245858;
   W_g[10,12] := 0.00857112;
   W_g[10,13] := 0.1074988;
   W_g[10,14] := -0.1275509;
   W_g[10,15] := -0.03629598;
   W_g[10,16] := -0.01334849;
   W_g[10,17] := 0.1290663;
   W_g[10,18] := -0.01503343;
   W_g[10,19] := 0.01173486;
   W_g[10,20] := 0.06222534;
   W_g[10,21] := 0.05678142;
   W_g[10,22] := -0.02349397;
   W_g[10,23] := 0.06754656;
   W_g[10,24] := 0.1779617;
   W_g[10,25] := 0.1916296;
   W_g[10,26] := -0.02255434;
   W_g[10,27] := 0.1007323;
   W_g[10,28] := 0.1328024;
   W_g[10,29] := -0.01282987;
   W_g[10,30] := -0.01621767;
   W_g[10,31] := -0.0140665;
   W_g[10,32] := -0.00099214;
   W_g[10,33] := -0.00035058;
   W_g[10,34] := 0.1452188;
   W_g[10,35] := 0.02793738;
   W_g[10,36] := -0.07625148;
   W_g[10,37] := -0.00763791;
   W_g[10,38] := 0.00534324;
   W_g[10,39] := -0.3312542;
   W_g[11,0] := -0.1137508;
   W_g[11,1] := 0.05398307;
   W_g[11,2] := -0.1207509;
   W_g[11,3] := 0.04525032;
   W_g[11,4] := 0.08992387;
   W_g[11,5] := 0.01991016;
   W_g[11,6] := 0.2249754;
   W_g[11,7] := 0.04191377;
   W_g[11,8] := 0.04533296;
   W_g[11,9] := 0.0449999;
   W_g[11,10] := -0.1099455;
   W_g[11,11] := 0.00437518;
   W_g[11,12] := -0.00140931;
   W_g[11,13] := 0.04130397;
   W_g[11,14] := 0.053694;
   W_g[11,15] := -0.00366092;
   W_g[11,16] := -0.07105832;
   W_g[11,17] := -0.07482163;
   W_g[11,18] := -0.07100122;
   W_g[11,19] := 0.01718117;
   W_g[11,20] := -0.1375782;
   W_g[11,21] := 0.113075;
   W_g[11,22] := 0.054169;
   W_g[11,23] := 0.02884634;
   W_g[11,24] := 0.5307817;
   W_g[11,25] := 0.3570411;
   W_g[11,26] := 0.03378;
   W_g[11,27] := 0.1037555;
   W_g[11,28] := 0.2505002;
   W_g[11,29] := -0.1244629;
   W_g[11,30] := 0.0558193;
   W_g[11,31] := 0.05851344;
   W_g[11,32] := 0.07730477;
   W_g[11,33] := 0.09541148;
   W_g[11,34] := 0.1203315;
   W_g[11,35] := 0.1210543;
   W_g[11,36] := -0.1949756;
   W_g[11,37] := 0.0137196;
   W_g[11,38] := 0.08832928;
   W_g[11,39] := 0.08146589;
   W_g[12,0] := -0.02631861;
   W_g[12,1] := 0.04126604;
   W_g[12,2] := -0.02663527;
   W_g[12,3] := -0.02984582;
   W_g[12,4] := -0.02636349;
   W_g[12,5] := 0.07986053;
   W_g[12,6] := -0.01390989;
   W_g[12,7] := -0.00909171;
   W_g[12,8] := -0.01941176;
   W_g[12,9] := -0.02868326;
   W_g[12,10] := 0.03089914;
   W_g[12,11] := 0.00787742;
   W_g[12,12] := -0.00904082;
   W_g[12,13] := -0.0291048;
   W_g[12,14] := 0.1083951;
   W_g[12,15] := 0.01380038;
   W_g[12,16] := 0.06520407;
   W_g[12,17] := -0.04494612;
   W_g[12,18] := -0.0019409;
   W_g[12,19] := -0.0150968;
   W_g[12,20] := 0.08029543;
   W_g[12,21] := 0.02437602;
   W_g[12,22] := -0.07042312;
   W_g[12,23] := -0.04948704;
   W_g[12,24] := -0.8303994;
   W_g[12,25] := -0.5589937;
   W_g[12,26] := -0.04566456;
   W_g[12,27] := 0.0018911;
   W_g[12,28] := -0.02951618;
   W_g[12,29] := -0.05513477;
   W_g[12,30] := -0.04795056;
   W_g[12,31] := -0.0368838;
   W_g[12,32] := -0.03588131;
   W_g[12,33] := 0.00737297;
   W_g[12,34] := 0.0499457;
   W_g[12,35] := -0.01839683;
   W_g[12,36] := -0.4987357;
   W_g[12,37] := -0.07791845;
   W_g[12,38] := -0.1047491;
   W_g[12,39] := 0.00553967;
   W_g[13,0] := -0.0268404;
   W_g[13,1] := -0.088905;
   W_g[13,2] := -0.02790045;
   W_g[13,3] := 0.08189317;
   W_g[13,4] := -0.1255152;
   W_g[13,5] := -0.05772218;
   W_g[13,6] := 0.09080454;
   W_g[13,7] := 0.08241173;
   W_g[13,8] := 0.07553043;
   W_g[13,9] := 0.08949121;
   W_g[13,10] := -0.02704351;
   W_g[13,11] := 0.00487661;
   W_g[13,12] := 0.02095871;
   W_g[13,13] := 0.06879441;
   W_g[13,14] := 0.00018557;
   W_g[13,15] := 0.01617457;
   W_g[13,16] := 0.2304675;
   W_g[13,17] := 0.08005539;
   W_g[13,18] := -0.06847396;
   W_g[13,19] := 0.02106568;
   W_g[13,20] := -0.08102658;
   W_g[13,21] := -0.03850572;
   W_g[13,22] := 0.00878646;
   W_g[13,23] := 0.1475209;
   W_g[13,24] := 0.1967756;
   W_g[13,25] := -0.00969006;
   W_g[13,26] := 0.04820746;
   W_g[13,27] := -0.06298333;
   W_g[13,28] := -0.06368192;
   W_g[13,29] := 0.01809042;
   W_g[13,30] := 0.01814866;
   W_g[13,31] := 0.00847225;
   W_g[13,32] := 0.00546922;
   W_g[13,33] := -0.01145526;
   W_g[13,34] := 0.1381362;
   W_g[13,35] := 0.01473064;
   W_g[13,36] := -0.050091;
   W_g[13,37] := -0.01566363;
   W_g[13,38] := 0.05946118;
   W_g[13,39] := 0.00826691;
   W_g[14,0] := 0.02104861;
   W_g[14,1] := 0.02198478;
   W_g[14,2] := 0.0111862;
   W_g[14,3] := -0.06436396;
   W_g[14,4] := 0.00489476;
   W_g[14,5] := 0.09250024;
   W_g[14,6] := -0.03399736;
   W_g[14,7] := -0.0496763;
   W_g[14,8] := -0.05370576;
   W_g[14,9] := -0.05536002;
   W_g[14,10] := 0.01229766;
   W_g[14,11] := -0.01784988;
   W_g[14,12] := -0.03607991;
   W_g[14,13] := 0.1900748;
   W_g[14,14] := 0.08048796;
   W_g[14,15] := -0.0089345;
   W_g[14,16] := 0.01208448;
   W_g[14,17] := -0.06566814;
   W_g[14,18] := -0.2211387;
   W_g[14,19] := -0.04166633;
   W_g[14,20] := 0.07567322;
   W_g[14,21] := -0.00166608;
   W_g[14,22] := -0.01256561;
   W_g[14,23] := 0.1539435;
   W_g[14,24] := 0.03526039;
   W_g[14,25] := 0.4811959;
   W_g[14,26] := 0.01489335;
   W_g[14,27] := 0.0317387;
   W_g[14,28] := 0.01991428;
   W_g[14,29] := 0.03107417;
   W_g[14,30] := -0.00682632;
   W_g[14,31] := 0.00660902;
   W_g[14,32] := 0.00283587;
   W_g[14,33] := -0.00859028;
   W_g[14,34] := -0.02930867;
   W_g[14,35] := 0.03631073;
   W_g[14,36] := 0.00467363;
   W_g[14,37] := 0.02703222;
   W_g[14,38] := -0.04237745;
   W_g[14,39] := 0.01309555;
   W_g[15,0] := 0.08495549;
   W_g[15,1] := -0.2072809;
   W_g[15,2] := 0.08629236;
   W_g[15,3] := -0.06330224;
   W_g[15,4] := 0.1923753;
   W_g[15,5] := 0.00801008;
   W_g[15,6] := -0.104994;
   W_g[15,7] := -0.05814644;
   W_g[15,8] := -0.06757385;
   W_g[15,9] := -0.0590176;
   W_g[15,10] := -0.00683508;
   W_g[15,11] := -0.00540838;
   W_g[15,12] := -0.02551957;
   W_g[15,13] := -0.01507952;
   W_g[15,14] := 0.00483655;
   W_g[15,15] := 0.01358667;
   W_g[15,16] := 0.2541837;
   W_g[15,17] := -0.01636837;
   W_g[15,18] := 0.01947031;
   W_g[15,19] := -0.03640394;
   W_g[15,20] := 0.2146612;
   W_g[15,21] := 0.1069127;
   W_g[15,22] := 0.03332973;
   W_g[15,23] := -0.06589723;
   W_g[15,24] := 0.1503799;
   W_g[15,25] := 0.03056319;
   W_g[15,26] := -0.08210966;
   W_g[15,27] := 0.1496714;
   W_g[15,28] := 0.09097399;
   W_g[15,29] := -0.04645663;
   W_g[15,30] := 0.04627259;
   W_g[15,31] := 0.00594573;
   W_g[15,32] := 0.05130993;
   W_g[15,33] := 0.05626767;
   W_g[15,34] := -0.00315162;
   W_g[15,35] := 0.04370028;
   W_g[15,36] := -0.06999733;
   W_g[15,37] := 0.01681984;
   W_g[15,38] := 0.0727107;
   W_g[15,39] := 0.01082875;
   W_o[0,0] := -0.1923357;
   W_o[0,1] := 0.1622824;
   W_o[0,2] := 0.03764162;
   W_o[0,3] := -0.00444271;
   W_o[0,4] := 0.0897337;
   W_o[0,5] := 0.05718408;
   W_o[0,6] := -0.2313943;
   W_o[0,7] := 0.1578357;
   W_o[0,8] := -0.1582883;
   W_o[0,9] := 0.1973625;
   W_o[0,10] := -0.3052712;
   W_o[0,11] := -0.2301492;
   W_o[0,12] := 0.209668;
   W_o[0,13] := -0.1742153;
   W_o[0,14] := -0.2678694;
   W_o[0,15] := -0.01321167;
   W_o[0,16] := -0.01970488;
   W_o[0,17] := -0.2028062;
   W_o[0,18] := 0.4272551;
   W_o[0,19] := -0.06582518;
   W_o[0,20] := -0.03046696;
   W_o[0,21] := 0.5501582;
   W_o[0,22] := 0.4423466;
   W_o[0,23] := -0.3345911;
   W_o[0,24] := 1.265247;
   W_o[0,25] := 1.416652;
   W_o[0,26] := -0.3267373;
   W_o[0,27] := -0.1832035;
   W_o[0,28] := 0.01126313;
   W_o[0,29] := -0.2838583;
   W_o[0,30] := 0.2609881;
   W_o[0,31] := 0.04669111;
   W_o[0,32] := 0.1043487;
   W_o[0,33] := 0.05575988;
   W_o[0,34] := 1.332353;
   W_o[0,35] := -0.06145113;
   W_o[0,36] := -0.0334513;
   W_o[0,37] := -0.2221547;
   W_o[0,38] := 0.00487359;
   W_o[0,39] := -0.03890218;
   W_o[1,0] := 0.7437804;
   W_o[1,1] := -0.0500013;
   W_o[1,2] := 0.1212982;
   W_o[1,3] := 0.1032013;
   W_o[1,4] := 0.1199842;
   W_o[1,5] := -0.1907221;
   W_o[1,6] := 0.2100161;
   W_o[1,7] := 0.1133247;
   W_o[1,8] := 0.3588262;
   W_o[1,9] := 0.3857575;
   W_o[1,10] := -0.4587842;
   W_o[1,11] := -0.1574819;
   W_o[1,12] := 0.2066407;
   W_o[1,13] := 0.1230617;
   W_o[1,14] := -0.203037;
   W_o[1,15] := 0.03768912;
   W_o[1,16] := -0.05619529;
   W_o[1,17] := -0.09439399;
   W_o[1,18] := 0.2707254;
   W_o[1,19] := 0.3822214;
   W_o[1,20] := -0.2934351;
   W_o[1,21] := 0.5161377;
   W_o[1,22] := 0.1759103;
   W_o[1,23] := 0.1837359;
   W_o[1,24] := -0.03005522;
   W_o[1,25] := 0.00781888;
   W_o[1,26] := -0.1068488;
   W_o[1,27] := -0.07173182;
   W_o[1,28] := 0.2014527;
   W_o[1,29] := 0.1306461;
   W_o[1,30] := -0.01024106;
   W_o[1,31] := -0.0716324;
   W_o[1,32] := 0.05804014;
   W_o[1,33] := 0.2721744;
   W_o[1,34] := 0.06194695;
   W_o[1,35] := -0.304073;
   W_o[1,36] := 0.1530892;
   W_o[1,37] := -0.07396729;
   W_o[1,38] := 0.08739793;
   W_o[1,39] := 0.3265531;
   W_o[2,0] := -0.03605163;
   W_o[2,1] := 0.07661975;
   W_o[2,2] := 0.1369504;
   W_o[2,3] := 0.09188601;
   W_o[2,4] := 0.03664814;
   W_o[2,5] := -0.02675835;
   W_o[2,6] := -0.01984608;
   W_o[2,7] := -0.1901468;
   W_o[2,8] := -0.02938575;
   W_o[2,9] := 0.1836661;
   W_o[2,10] := -0.1862541;
   W_o[2,11] := 0.06671655;
   W_o[2,12] := 0.3190728;
   W_o[2,13] := -0.01547686;
   W_o[2,14] := -0.05195596;
   W_o[2,15] := 0.03504787;
   W_o[2,16] := 0.3541903;
   W_o[2,17] := 0.02718459;
   W_o[2,18] := -0.2491126;
   W_o[2,19] := -0.8667619;
   W_o[2,20] := -0.1266757;
   W_o[2,21] := 0.02015731;
   W_o[2,22] := -0.02294585;
   W_o[2,23] := -0.01648583;
   W_o[2,24] := -0.1919154;
   W_o[2,25] := 0.00051678;
   W_o[2,26] := 0.06543333;
   W_o[2,27] := 0.1037415;
   W_o[2,28] := -0.0450457;
   W_o[2,29] := 0.215062;
   W_o[2,30] := 0.02658869;
   W_o[2,31] := -0.1369152;
   W_o[2,32] := 0.01719045;
   W_o[2,33] := 0.218743;
   W_o[2,34] := -0.07076459;
   W_o[2,35] := -0.0740788;
   W_o[2,36] := -0.08052358;
   W_o[2,37] := -0.2012888;
   W_o[2,38] := -0.3849033;
   W_o[2,39] := 0.6891636;
   W_o[3,0] := -0.06302688;
   W_o[3,1] := 0.2002212;
   W_o[3,2] := 0.0159587;
   W_o[3,3] := -0.0018361;
   W_o[3,4] := -0.8591735;
   W_o[3,5] := 0.1731812;
   W_o[3,6] := 0.2409841;
   W_o[3,7] := 0.2596082;
   W_o[3,8] := -0.00940404;
   W_o[3,9] := 0.06814823;
   W_o[3,10] := -0.01664601;
   W_o[3,11] := 0.148778;
   W_o[3,12] := -0.09583785;
   W_o[3,13] := -0.2798349;
   W_o[3,14] := 0.1443422;
   W_o[3,15] := 0.00555357;
   W_o[3,16] := -0.02839783;
   W_o[3,17] := 0.09947813;
   W_o[3,18] := 0.4643263;
   W_o[3,19] := 0.0636435;
   W_o[3,20] := -0.08531965;
   W_o[3,21] := 1.165775;
   W_o[3,22] := 0.3448276;
   W_o[3,23] := -0.117277;
   W_o[3,24] := 1.352477;
   W_o[3,25] := 1.178241;
   W_o[3,26] := -0.4892529;
   W_o[3,27] := -0.7737502;
   W_o[3,28] := 0.2264518;
   W_o[3,29] := 0.00574818;
   W_o[3,30] := 0.2461463;
   W_o[3,31] := 0.1052826;
   W_o[3,32] := 0.00088265;
   W_o[3,33] := 0.1049805;
   W_o[3,34] := 1.18573;
   W_o[3,35] := 0.1909419;
   W_o[3,36] := -0.00811989;
   W_o[3,37] := 0.09236411;
   W_o[3,38] := 0.1108437;
   W_o[3,39] := 0.9237891;
   W_o[4,0] := -0.1855668;
   W_o[4,1] := -0.06182796;
   W_o[4,2] := 0.1497869;
   W_o[4,3] := -0.02874054;
   W_o[4,4] := -0.2372189;
   W_o[4,5] := -0.02661614;
   W_o[4,6] := 0.04865195;
   W_o[4,7] := -0.2595509;
   W_o[4,8] := 0.5146528;
   W_o[4,9] := -0.2822051;
   W_o[4,10] := 0.01177313;
   W_o[4,11] := -0.4989094;
   W_o[4,12] := -0.8648744;
   W_o[4,13] := -0.04488994;
   W_o[4,14] := -0.0542339;
   W_o[4,15] := -0.5589076;
   W_o[4,16] := -0.145594;
   W_o[4,17] := 0.02167914;
   W_o[4,18] := 1.006644;
   W_o[4,19] := -0.2599575;
   W_o[4,20] := 0.00703312;
   W_o[4,21] := -0.2283233;
   W_o[4,22] := 0.00192229;
   W_o[4,23] := -0.01435418;
   W_o[4,24] := 0.04472705;
   W_o[4,25] := 0.2338529;
   W_o[4,26] := -0.1127145;
   W_o[4,27] := 0.08130027;
   W_o[4,28] := 0.4603895;
   W_o[4,29] := 0.1379606;
   W_o[4,30] := 0.1812189;
   W_o[4,31] := -0.3901244;
   W_o[4,32] := -0.0703788;
   W_o[4,33] := 0.2888122;
   W_o[4,34] := 0.4034505;
   W_o[4,35] := 0.0328819;
   W_o[4,36] := -0.09105004;
   W_o[4,37] := 0.09711539;
   W_o[4,38] := -0.1910721;
   W_o[4,39] := -0.01934181;
   W_o[5,0] := -0.6595194;
   W_o[5,1] := 0.3772199;
   W_o[5,2] := 0.00501744;
   W_o[5,3] := 0.532542;
   W_o[5,4] := 0.2366183;
   W_o[5,5] := 1.09201;
   W_o[5,6] := 0.9502543;
   W_o[5,7] := 0.2582511;
   W_o[5,8] := -0.4691281;
   W_o[5,9] := 0.3928114;
   W_o[5,10] := 1.11464;
   W_o[5,11] := -0.7781826;
   W_o[5,12] := -0.6074764;
   W_o[5,13] := 0.16801;
   W_o[5,14] := -0.1086531;
   W_o[5,15] := -0.6841738;
   W_o[5,16] := -0.3678641;
   W_o[5,17] := -0.2172338;
   W_o[5,18] := 0.3863191;
   W_o[5,19] := -0.4950597;
   W_o[5,20] := -0.5119882;
   W_o[5,21] := -0.1780492;
   W_o[5,22] := 0.1544936;
   W_o[5,23] := 0.1383117;
   W_o[5,24] := 1.004889;
   W_o[5,25] := 1.139415;
   W_o[5,26] := -0.3015366;
   W_o[5,27] := -0.04238907;
   W_o[5,28] := -0.3108428;
   W_o[5,29] := 0.3969988;
   W_o[5,30] := 0.01171695;
   W_o[5,31] := -0.3139689;
   W_o[5,32] := -0.3243381;
   W_o[5,33] := -0.414901;
   W_o[5,34] := 0.2215569;
   W_o[5,35] := -0.133694;
   W_o[5,36] := 0.02332771;
   W_o[5,37] := -0.1487403;
   W_o[5,38] := 0.1979396;
   W_o[5,39] := -0.2030152;
   W_o[6,0] := -0.04529256;
   W_o[6,1] := 0.2150283;
   W_o[6,2] := 0.09295318;
   W_o[6,3] := -0.0767066;
   W_o[6,4] := -0.1236452;
   W_o[6,5] := 0.3573766;
   W_o[6,6] := -0.2646887;
   W_o[6,7] := 0.2834802;
   W_o[6,8] := -0.04882327;
   W_o[6,9] := 0.8413;
   W_o[6,10] := 1.089968;
   W_o[6,11] := -0.06981075;
   W_o[6,12] := 0.05921048;
   W_o[6,13] := -0.5099319;
   W_o[6,14] := 0.04131682;
   W_o[6,15] := 0.09513918;
   W_o[6,16] := 0.08072844;
   W_o[6,17] := 0.02096614;
   W_o[6,18] := 0.1683812;
   W_o[6,19] := 0.1104724;
   W_o[6,20] := -0.3392214;
   W_o[6,21] := -0.09979945;
   W_o[6,22] := 0.1501902;
   W_o[6,23] := -0.06504018;
   W_o[6,24] := 1.949389;
   W_o[6,25] := 1.979982;
   W_o[6,26] := 0.02307883;
   W_o[6,27] := 0.2684888;
   W_o[6,28] := 0.09674384;
   W_o[6,29] := 0.2116341;
   W_o[6,30] := 0.1413678;
   W_o[6,31] := -0.0124489;
   W_o[6,32] := -0.04519035;
   W_o[6,33] := -0.1396772;
   W_o[6,34] := 0.4939206;
   W_o[6,35] := -0.2130735;
   W_o[6,36] := 0.06053885;
   W_o[6,37] := 0.0587407;
   W_o[6,38] := 0.429702;
   W_o[6,39] := -0.1062183;
   W_o[7,0] := 0.1648133;
   W_o[7,1] := -0.09838933;
   W_o[7,2] := -0.0939215;
   W_o[7,3] := -0.1272545;
   W_o[7,4] := -0.2333547;
   W_o[7,5] := 0.05955706;
   W_o[7,6] := 0.2717095;
   W_o[7,7] := 0.1100897;
   W_o[7,8] := 0.1809682;
   W_o[7,9] := 0.01596895;
   W_o[7,10] := 0.1498611;
   W_o[7,11] := -0.3100757;
   W_o[7,12] := 0.5308929;
   W_o[7,13] := -0.07378945;
   W_o[7,14] := -0.2509805;
   W_o[7,15] := 0.2649329;
   W_o[7,16] := -0.1476106;
   W_o[7,17] := -0.2392291;
   W_o[7,18] := 0.4080176;
   W_o[7,19] := -0.1504776;
   W_o[7,20] := -0.1111432;
   W_o[7,21] := 0.1132136;
   W_o[7,22] := 0.464526;
   W_o[7,23] := -0.1314203;
   W_o[7,24] := 0.8524858;
   W_o[7,25] := 0.9319458;
   W_o[7,26] := 0.1910378;
   W_o[7,27] := -0.04179411;
   W_o[7,28] := 0.1727818;
   W_o[7,29] := -0.3418947;
   W_o[7,30] := 0.4730469;
   W_o[7,31] := 0.08789608;
   W_o[7,32] := 0.2170709;
   W_o[7,33] := -0.03279238;
   W_o[7,34] := 0.6582685;
   W_o[7,35] := 0.08038806;
   W_o[7,36] := 0.04812925;
   W_o[7,37] := 0.4378351;
   W_o[7,38] := -0.06570955;
   W_o[7,39] := -1.681702;
   W_o[8,0] := 0.2838559;
   W_o[8,1] := -0.1376109;
   W_o[8,2] := -0.00303996;
   W_o[8,3] := -0.1514946;
   W_o[8,4] := -0.05367951;
   W_o[8,5] := 0.3758456;
   W_o[8,6] := 0.02626968;
   W_o[8,7] := -0.1422179;
   W_o[8,8] := 0.00944922;
   W_o[8,9] := -0.2079319;
   W_o[8,10] := -0.2131251;
   W_o[8,11] := -1.025984;
   W_o[8,12] := -0.3985277;
   W_o[8,13] := -0.0818603;
   W_o[8,14] := -0.1052002;
   W_o[8,15] := -1.120577;
   W_o[8,16] := 0.05219958;
   W_o[8,17] := 0.7909105;
   W_o[8,18] := 0.3779635;
   W_o[8,19] := 0.16329;
   W_o[8,20] := -0.06752818;
   W_o[8,21] := 0.2244961;
   W_o[8,22] := -0.133298;
   W_o[8,23] := -0.5498607;
   W_o[8,24] := 0.210675;
   W_o[8,25] := 0.4249826;
   W_o[8,26] := 0.3085507;
   W_o[8,27] := 0.00327513;
   W_o[8,28] := -0.1328674;
   W_o[8,29] := 0.2423343;
   W_o[8,30] := -0.2916745;
   W_o[8,31] := 0.1113145;
   W_o[8,32] := 0.235408;
   W_o[8,33] := 0.2593887;
   W_o[8,34] := 0.2619374;
   W_o[8,35] := 0.09260385;
   W_o[8,36] := -0.07284077;
   W_o[8,37] := 0.2716717;
   W_o[8,38] := -0.5921684;
   W_o[8,39] := 0.1613293;
   W_o[9,0] := -0.6345086;
   W_o[9,1] := -0.259372;
   W_o[9,2] := -0.4410478;
   W_o[9,3] := -0.1479532;
   W_o[9,4] := 0.07470662;
   W_o[9,5] := -0.1442392;
   W_o[9,6] := 0.2044672;
   W_o[9,7] := -0.3629733;
   W_o[9,8] := -0.8357224;
   W_o[9,9] := -0.03687909;
   W_o[9,10] := -0.5277801;
   W_o[9,11] := 0.1395604;
   W_o[9,12] := 0.00705423;
   W_o[9,13] := -0.06065191;
   W_o[9,14] := 0.00270301;
   W_o[9,15] := 0.02473978;
   W_o[9,16] := -0.1366292;
   W_o[9,17] := -0.1191437;
   W_o[9,18] := -0.06459489;
   W_o[9,19] := -0.155962;
   W_o[9,20] := -0.1332201;
   W_o[9,21] := 0.6168138;
   W_o[9,22] := -0.008209;
   W_o[9,23] := -0.03221058;
   W_o[9,24] := -0.07914114;
   W_o[9,25] := -0.2822376;
   W_o[9,26] := 0.1799158;
   W_o[9,27] := 0.1354283;
   W_o[9,28] := 0.1905717;
   W_o[9,29] := 0.3257442;
   W_o[9,30] := 0.2045423;
   W_o[9,31] := 0.117547;
   W_o[9,32] := 0.1869259;
   W_o[9,33] := 0.4169515;
   W_o[9,34] := 0.131826;
   W_o[9,35] := -0.1867882;
   W_o[9,36] := -0.09728058;
   W_o[9,37] := -0.2151765;
   W_o[9,38] := 0.03850761;
   W_o[9,39] := -0.0044641;
   W_o[10,0] := 0.06105608;
   W_o[10,1] := -0.06832715;
   W_o[10,2] := 0.07474305;
   W_o[10,3] := -0.08913961;
   W_o[10,4] := -0.2327598;
   W_o[10,5] := 0.07582341;
   W_o[10,6] := 0.104368;
   W_o[10,7] := 0.03688281;
   W_o[10,8] := -0.01102509;
   W_o[10,9] := -0.02805536;
   W_o[10,10] := 0.1092547;
   W_o[10,11] := -0.04491638;
   W_o[10,12] := -0.00955069;
   W_o[10,13] := -0.3600228;
   W_o[10,14] := -0.2598117;
   W_o[10,15] := -0.1312952;
   W_o[10,16] := 0.1270282;
   W_o[10,17] := 0.2455932;
   W_o[10,18] := 0.02347365;
   W_o[10,19] := 0.08953306;
   W_o[10,20] := -0.412829;
   W_o[10,21] := -0.1269261;
   W_o[10,22] := 0.1430949;
   W_o[10,23] := -0.2883692;
   W_o[10,24] := 1.613103;
   W_o[10,25] := 1.56905;
   W_o[10,26] := 0.11707;
   W_o[10,27] := -0.6253218;
   W_o[10,28] := -0.570655;
   W_o[10,29] := 0.06348585;
   W_o[10,30] := 0.2199306;
   W_o[10,31] := -0.02762064;
   W_o[10,32] := 0.08508236;
   W_o[10,33] := 0.2603731;
   W_o[10,34] := 0.5238683;
   W_o[10,35] := -0.3072915;
   W_o[10,36] := 0.4589803;
   W_o[10,37] := -0.3261147;
   W_o[10,38] := -0.04951124;
   W_o[10,39] := -0.0165583;
   W_o[11,0] := 0.2717895;
   W_o[11,1] := 0.4973186;
   W_o[11,2] := -0.111147;
   W_o[11,3] := 0.00516717;
   W_o[11,4] := -0.7287747;
   W_o[11,5] := -0.07876529;
   W_o[11,6] := -0.5072603;
   W_o[11,7] := -0.03536538;
   W_o[11,8] := 0.1201321;
   W_o[11,9] := 0.1112787;
   W_o[11,10] := 0.1532365;
   W_o[11,11] := -0.4891608;
   W_o[11,12] := 0.1887655;
   W_o[11,13] := 0.1852349;
   W_o[11,14] := 0.1703349;
   W_o[11,15] := -0.2467272;
   W_o[11,16] := 0.04845995;
   W_o[11,17] := 0.2819173;
   W_o[11,18] := 0.1057306;
   W_o[11,19] := -0.00306271;
   W_o[11,20] := -0.724054;
   W_o[11,21] := 0.09254762;
   W_o[11,22] := -0.4099866;
   W_o[11,23] := -0.1073627;
   W_o[11,24] := -0.0586772;
   W_o[11,25] := 0.3430104;
   W_o[11,26] := 0.1855343;
   W_o[11,27] := 0.1084731;
   W_o[11,28] := 0.5040212;
   W_o[11,29] := -0.00853192;
   W_o[11,30] := -0.3662441;
   W_o[11,31] := -0.01966033;
   W_o[11,32] := -0.06275205;
   W_o[11,33] := 0.09751767;
   W_o[11,34] := -0.2004695;
   W_o[11,35] := -0.1034404;
   W_o[11,36] := 0.2302412;
   W_o[11,37] := 0.1414506;
   W_o[11,38] := 0.266502;
   W_o[11,39] := -0.3097887;
   W_o[12,0] := -0.01830707;
   W_o[12,1] := 0.131161;
   W_o[12,2] := 0.00496979;
   W_o[12,3] := 0.2061931;
   W_o[12,4] := 0.03057155;
   W_o[12,5] := 0.02297443;
   W_o[12,6] := 0.05931674;
   W_o[12,7] := -0.03210922;
   W_o[12,8] := 0.07573608;
   W_o[12,9] := 0.1248056;
   W_o[12,10] := -0.07253183;
   W_o[12,11] := -0.2442229;
   W_o[12,12] := 0.1326389;
   W_o[12,13] := -0.1664325;
   W_o[12,14] := -0.1405273;
   W_o[12,15] := -0.05658006;
   W_o[12,16] := 0.04406866;
   W_o[12,17] := 0.0236842;
   W_o[12,18] := 0.7910394;
   W_o[12,19] := 0.02559086;
   W_o[12,20] := -0.1635535;
   W_o[12,21] := -0.01013497;
   W_o[12,22] := -0.3506611;
   W_o[12,23] := -0.1885774;
   W_o[12,24] := 0.4997112;
   W_o[12,25] := 0.5154855;
   W_o[12,26] := 0.1843938;
   W_o[12,27] := 0.02656424;
   W_o[12,28] := 0.00674596;
   W_o[12,29] := 0.03458697;
   W_o[12,30] := -0.4318717;
   W_o[12,31] := -0.1312484;
   W_o[12,32] := -0.3812101;
   W_o[12,33] := -0.02800291;
   W_o[12,34] := -0.2285903;
   W_o[12,35] := 0.123769;
   W_o[12,36] := 0.08067092;
   W_o[12,37] := -0.04127869;
   W_o[12,38] := -0.06010977;
   W_o[12,39] := -0.00181283;
   W_o[13,0] := -0.04045204;
   W_o[13,1] := -0.3968439;
   W_o[13,2] := 0.08165251;
   W_o[13,3] := -0.01278869;
   W_o[13,4] := -0.4479226;
   W_o[13,5] := -0.2656083;
   W_o[13,6] := 0.3235124;
   W_o[13,7] := 0.574206;
   W_o[13,8] := -0.2794143;
   W_o[13,9] := 0.3598377;
   W_o[13,10] := -0.08126416;
   W_o[13,11] := -0.00919488;
   W_o[13,12] := 0.09122144;
   W_o[13,13] := 0.02155786;
   W_o[13,14] := 0.1209246;
   W_o[13,15] := -0.00289959;
   W_o[13,16] := -0.2549352;
   W_o[13,17] := -0.2486969;
   W_o[13,18] := 0.6917394;
   W_o[13,19] := -0.03206153;
   W_o[13,20] := -0.2219304;
   W_o[13,21] := 0.1183459;
   W_o[13,22] := 0.3679306;
   W_o[13,23] := 0.4413242;
   W_o[13,24] := 1.975207;
   W_o[13,25] := 1.843769;
   W_o[13,26] := -0.279261;
   W_o[13,27] := -0.3077843;
   W_o[13,28] := -0.01960251;
   W_o[13,29] := -0.2369677;
   W_o[13,30] := 0.109645;
   W_o[13,31] := -0.1079782;
   W_o[13,32] := 0.038799;
   W_o[13,33] := 0.05485996;
   W_o[13,34] := 0.5972548;
   W_o[13,35] := 0.01886969;
   W_o[13,36] := 0.09835773;
   W_o[13,37] := 0.3843534;
   W_o[13,38] := 0.05617079;
   W_o[13,39] := -0.2227704;
   W_o[14,0] := 0.8289077;
   W_o[14,1] := -0.2031105;
   W_o[14,2] := 0.03403382;
   W_o[14,3] := 0.05452057;
   W_o[14,4] := 0.2272833;
   W_o[14,5] := -0.07046781;
   W_o[14,6] := 0.3896516;
   W_o[14,7] := 0.4871905;
   W_o[14,8] := -0.07724485;
   W_o[14,9] := -0.07247894;
   W_o[14,10] := 0.2814783;
   W_o[14,11] := -0.02350411;
   W_o[14,12] := 0.3741138;
   W_o[14,13] := 0.01457606;
   W_o[14,14] := -0.08907567;
   W_o[14,15] := 0.03109477;
   W_o[14,16] := 0.05151353;
   W_o[14,17] := -0.1566754;
   W_o[14,18] := -0.2640311;
   W_o[14,19] := -0.1076154;
   W_o[14,20] := 0.3854151;
   W_o[14,21] := 1.575822;
   W_o[14,22] := -0.05344179;
   W_o[14,23] := -0.9402446;
   W_o[14,24] := -0.0189026;
   W_o[14,25] := -0.00721721;
   W_o[14,26] := -0.4206359;
   W_o[14,27] := 0.5079048;
   W_o[14,28] := 0.2300513;
   W_o[14,29] := 0.2341685;
   W_o[14,30] := -0.1072616;
   W_o[14,31] := -0.05015407;
   W_o[14,32] := 0.03626099;
   W_o[14,33] := 0.2209553;
   W_o[14,34] := 0.2829649;
   W_o[14,35] := -0.102007;
   W_o[14,36] := 0.00415739;
   W_o[14,37] := 0.2021578;
   W_o[14,38] := 0.1449325;
   W_o[14,39] := 0.1953939;
   W_o[15,0] := 0.00236452;
   W_o[15,1] := 0.6316325;
   W_o[15,2] := 0.04516845;
   W_o[15,3] := -0.1972448;
   W_o[15,4] := -0.6675987;
   W_o[15,5] := 0.3806524;
   W_o[15,6] := 0.6475521;
   W_o[15,7] := 0.2695197;
   W_o[15,8] := -0.4985425;
   W_o[15,9] := -0.3775528;
   W_o[15,10] := 0.255392;
   W_o[15,11] := -0.1499313;
   W_o[15,12] := 0.5755351;
   W_o[15,13] := -0.03951031;
   W_o[15,14] := 0.02471058;
   W_o[15,15] := -0.2347889;
   W_o[15,16] := 0.3119133;
   W_o[15,17] := 0.02724188;
   W_o[15,18] := 0.3374691;
   W_o[15,19] := -0.0329643;
   W_o[15,20] := -0.8862573;
   W_o[15,21] := 0.5019892;
   W_o[15,22] := -0.01491885;
   W_o[15,23] := 0.393534;
   W_o[15,24] := 0.2951014;
   W_o[15,25] := 0.4423684;
   W_o[15,26] := -0.03397221;
   W_o[15,27] := -0.4513796;
   W_o[15,28] := 0.261473;
   W_o[15,29] := -0.1054694;
   W_o[15,30] := 0.3078526;
   W_o[15,31] := -0.1044204;
   W_o[15,32] := 0.2778185;
   W_o[15,33] := -0.00624027;
   W_o[15,34] := 0.2965292;
   W_o[15,35] := -0.2159247;
   W_o[15,36] := 0.05058118;
   W_o[15,37] := 0.00013962;
   W_o[15,38] := 1.000757;
   W_o[15,39] := 0.5571635;
   R_i[0,0] := -0.1137149;
   R_i[0,1] := -0.00305563;
   R_i[0,2] := 0.4498252;
   R_i[0,3] := 0.408096;
   R_i[0,4] := 0.4966823;
   R_i[0,5] := 0.2685225;
   R_i[0,6] := 0.5829936;
   R_i[0,7] := 0.309512;
   R_i[0,8] := 0.584756;
   R_i[0,9] := 0.4425567;
   R_i[0,10] := 0.168636;
   R_i[0,11] := -0.314454;
   R_i[0,12] := 0.01961905;
   R_i[0,13] := 0.3972826;
   R_i[0,14] := 0.3588874;
   R_i[0,15] := 0.1209446;
   R_i[1,0] := -0.03926941;
   R_i[1,1] := -0.2256729;
   R_i[1,2] := -0.1890858;
   R_i[1,3] := -0.4077013;
   R_i[1,4] := 1.580356;
   R_i[1,5] := -0.5334294;
   R_i[1,6] := -0.07024953;
   R_i[1,7] := 0.4276721;
   R_i[1,8] := -0.6611474;
   R_i[1,9] := 0.4677508;
   R_i[1,10] := -0.07782394;
   R_i[1,11] := -0.4426747;
   R_i[1,12] := 0.1923219;
   R_i[1,13] := 0.6306989;
   R_i[1,14] := -0.442345;
   R_i[1,15] := -0.1436543;
   R_i[2,0] := -0.1087616;
   R_i[2,1] := -0.00270978;
   R_i[2,2] := 0.2189552;
   R_i[2,3] := -0.5836519;
   R_i[2,4] := -0.07285596;
   R_i[2,5] := 0.04414057;
   R_i[2,6] := 0.2944021;
   R_i[2,7] := -0.5636789;
   R_i[2,8] := 0.02525483;
   R_i[2,9] := 0.2138523;
   R_i[2,10] := 0.1495301;
   R_i[2,11] := 0.4767698;
   R_i[2,12] := 0.3593693;
   R_i[2,13] := -0.475326;
   R_i[2,14] := -0.06119934;
   R_i[2,15] := -0.1814424;
   R_i[3,0] := -0.3477732;
   R_i[3,1] := -0.02923841;
   R_i[3,2] := -0.01545414;
   R_i[3,3] := 0.6730511;
   R_i[3,4] := 0.5243366;
   R_i[3,5] := 0.1240829;
   R_i[3,6] := 0.3667154;
   R_i[3,7] := 0.4002697;
   R_i[3,8] := 0.66468;
   R_i[3,9] := 0.1677333;
   R_i[3,10] := 0.1911234;
   R_i[3,11] := -0.5108734;
   R_i[3,12] := 0.1124746;
   R_i[3,13] := -0.2656624;
   R_i[3,14] := 0.3824491;
   R_i[3,15] := -0.1521915;
   R_i[4,0] := 0.00580328;
   R_i[4,1] := 0.6645847;
   R_i[4,2] := -0.7531157;
   R_i[4,3] := 0.00536597;
   R_i[4,4] := -1.547926;
   R_i[4,5] := -0.4703412;
   R_i[4,6] := -0.2358381;
   R_i[4,7] := 0.2062922;
   R_i[4,8] := 0.5056434;
   R_i[4,9] := 0.1705665;
   R_i[4,10] := -0.126984;
   R_i[4,11] := -1.014073;
   R_i[4,12] := 0.5201921;
   R_i[4,13] := -0.1478145;
   R_i[4,14] := -0.1872073;
   R_i[4,15] := -0.01908887;
   R_i[5,0] := -0.5724422;
   R_i[5,1] := 0.07744113;
   R_i[5,2] := 0.07027231;
   R_i[5,3] := 0.1578984;
   R_i[5,4] := 0.2315233;
   R_i[5,5] := 0.1378991;
   R_i[5,6] := -0.3647587;
   R_i[5,7] := -0.1986962;
   R_i[5,8] := -0.04011904;
   R_i[5,9] := -0.05832585;
   R_i[5,10] := -0.04800356;
   R_i[5,11] := -0.2021917;
   R_i[5,12] := -0.02367323;
   R_i[5,13] := 0.1801978;
   R_i[5,14] := 0.07786623;
   R_i[5,15] := -0.4144403;
   R_i[6,0] := -0.4898062;
   R_i[6,1] := -0.08807379;
   R_i[6,2] := 0.729624;
   R_i[6,3] := 0.5344335;
   R_i[6,4] := -0.3394561;
   R_i[6,5] := 0.02468326;
   R_i[6,6] := -0.5965754;
   R_i[6,7] := -0.1523064;
   R_i[6,8] := -0.06543954;
   R_i[6,9] := 0.0652044;
   R_i[6,10] := -0.09473334;
   R_i[6,11] := 0.06633532;
   R_i[6,12] := 0.5554917;
   R_i[6,13] := -0.5657542;
   R_i[6,14] := 0.1251685;
   R_i[6,15] := -1.210496;
   R_i[7,0] := 0.09141196;
   R_i[7,1] := -0.2953948;
   R_i[7,2] := -0.04736479;
   R_i[7,3] := 0.6381459;
   R_i[7,4] := -0.1735898;
   R_i[7,5] := 0.02200026;
   R_i[7,6] := -0.542483;
   R_i[7,7] := 0.4112348;
   R_i[7,8] := 0.08935327;
   R_i[7,9] := 0.211784;
   R_i[7,10] := 0.3778164;
   R_i[7,11] := -0.2455601;
   R_i[7,12] := -0.2529224;
   R_i[7,13] := 0.3676308;
   R_i[7,14] := -0.1642352;
   R_i[7,15] := 0.3013193;
   R_i[8,0] := -0.4359751;
   R_i[8,1] := 0.5370886;
   R_i[8,2] := -0.01918638;
   R_i[8,3] := 0.06577428;
   R_i[8,4] := -0.2360706;
   R_i[8,5] := 0.04361986;
   R_i[8,6] := 0.4372621;
   R_i[8,7] := 0.317978;
   R_i[8,8] := -1.000937;
   R_i[8,9] := -0.3358858;
   R_i[8,10] := 0.9401911;
   R_i[8,11] := -0.4844143;
   R_i[8,12] := -0.02272851;
   R_i[8,13] := 0.1828933;
   R_i[8,14] := -0.01882748;
   R_i[8,15] := -0.06172743;
   R_i[9,0] := -0.5143862;
   R_i[9,1] := 0.06295519;
   R_i[9,2] := 0.3046114;
   R_i[9,3] := 0.03788998;
   R_i[9,4] := 0.1308033;
   R_i[9,5] := -0.358474;
   R_i[9,6] := 0.69233;
   R_i[9,7] := -0.2776851;
   R_i[9,8] := 0.00155199;
   R_i[9,9] := -0.09497612;
   R_i[9,10] := 0.191216;
   R_i[9,11] := -0.428836;
   R_i[9,12] := 0.097583;
   R_i[9,13] := 0.2892125;
   R_i[9,14] := 0.1341387;
   R_i[9,15] := -0.6526389;
   R_i[10,0] := -1.243925;
   R_i[10,1] := 0.680451;
   R_i[10,2] := 0.9452817;
   R_i[10,3] := -1.115271;
   R_i[10,4] := -0.6274545;
   R_i[10,5] := -0.4702299;
   R_i[10,6] := 0.9055709;
   R_i[10,7] := 0.7863802;
   R_i[10,8] := 1.259396;
   R_i[10,9] := 0.4866133;
   R_i[10,10] := -0.232237;
   R_i[10,11] := -0.8811347;
   R_i[10,12] := -0.1416707;
   R_i[10,13] := 0.2519798;
   R_i[10,14] := 0.7145844;
   R_i[10,15] := -0.03913529;
   R_i[11,0] := -0.2986307;
   R_i[11,1] := 0.7416621;
   R_i[11,2] := -0.5418634;
   R_i[11,3] := -0.0208676;
   R_i[11,4] := 0.4454969;
   R_i[11,5] := -0.1592286;
   R_i[11,6] := 0.2505509;
   R_i[11,7] := -0.382692;
   R_i[11,8] := 0.1618413;
   R_i[11,9] := 0.4193928;
   R_i[11,10] := 0.02712804;
   R_i[11,11] := -1.186852;
   R_i[11,12] := 0.2001949;
   R_i[11,13] := 0.1532502;
   R_i[11,14] := -0.3284004;
   R_i[11,15] := -0.2820552;
   R_i[12,0] := -0.2895075;
   R_i[12,1] := 1.091435;
   R_i[12,2] := -0.05338987;
   R_i[12,3] := 0.2911161;
   R_i[12,4] := 0.1629717;
   R_i[12,5] := -0.161591;
   R_i[12,6] := 0.5146877;
   R_i[12,7] := 0.03626299;
   R_i[12,8] := 0.08357667;
   R_i[12,9] := 0.2767582;
   R_i[12,10] := -0.2725959;
   R_i[12,11] := -0.9445232;
   R_i[12,12] := 2.164176;
   R_i[12,13] := -0.04564672;
   R_i[12,14] := -0.9437686;
   R_i[12,15] := -0.3752556;
   R_i[13,0] := -0.3738814;
   R_i[13,1] := -0.4302073;
   R_i[13,2] := 0.06173271;
   R_i[13,3] := -0.3280604;
   R_i[13,4] := -0.2716264;
   R_i[13,5] := 0.3550667;
   R_i[13,6] := -0.05685175;
   R_i[13,7] := 0.5135436;
   R_i[13,8] := 0.1640313;
   R_i[13,9] := -0.2691319;
   R_i[13,10] := -0.3801848;
   R_i[13,11] := 0.1228051;
   R_i[13,12] := 0.5428029;
   R_i[13,13] := 1.709359;
   R_i[13,14] := 1.011569;
   R_i[13,15] := -0.4288203;
   R_i[14,0] := 0.2300761;
   R_i[14,1] := -1.012092;
   R_i[14,2] := 0.6361403;
   R_i[14,3] := 0.05786986;
   R_i[14,4] := -0.4553789;
   R_i[14,5] := -0.6679262;
   R_i[14,6] := -0.4034081;
   R_i[14,7] := 0.00973069;
   R_i[14,8] := 1.011842;
   R_i[14,9] := -0.3590509;
   R_i[14,10] := 0.3335861;
   R_i[14,11] := -0.8217174;
   R_i[14,12] := -0.6475059;
   R_i[14,13] := -0.2020338;
   R_i[14,14] := 3.036138;
   R_i[14,15] := -0.1744984;
   R_i[15,0] := -0.04125203;
   R_i[15,1] := 0.6700256;
   R_i[15,2] := 1.07735;
   R_i[15,3] := 0.2874972;
   R_i[15,4] := -0.03804383;
   R_i[15,5] := 0.0777116;
   R_i[15,6] := 0.6422315;
   R_i[15,7] := 0.2854839;
   R_i[15,8] := 0.2419276;
   R_i[15,9] := 0.0058566;
   R_i[15,10] := 0.6288991;
   R_i[15,11] := -0.8346034;
   R_i[15,12] := 0.2495139;
   R_i[15,13] := -0.4616964;
   R_i[15,14] := 0.8547717;
   R_i[15,15] := -1.059702;
   R_f[0,0] := 0.3233714;
   R_f[0,1] := -0.6415426;
   R_f[0,2] := 0.4436696;
   R_f[0,3] := -0.1691184;
   R_f[0,4] := -0.2260693;
   R_f[0,5] := 0.4070715;
   R_f[0,6] := 0.9958715;
   R_f[0,7] := -0.6152283;
   R_f[0,8] := -0.1669062;
   R_f[0,9] := 0.1140058;
   R_f[0,10] := -1.301264;
   R_f[0,11] := 0.6843588;
   R_f[0,12] := 0.2550505;
   R_f[0,13] := -0.5000576;
   R_f[0,14] := 1.899208;
   R_f[0,15] := 0.3119706;
   R_f[1,0] := -0.1011617;
   R_f[1,1] := 3.477333;
   R_f[1,2] := -0.2395845;
   R_f[1,3] := 0.2576158;
   R_f[1,4] := 0.6485823;
   R_f[1,5] := 0.2552066;
   R_f[1,6] := 0.4734288;
   R_f[1,7] := 0.4439468;
   R_f[1,8] := 0.08832169;
   R_f[1,9] := -0.07672439;
   R_f[1,10] := -0.1136505;
   R_f[1,11] := -0.1276775;
   R_f[1,12] := 0.153016;
   R_f[1,13] := 0.1081575;
   R_f[1,14] := -0.00451868;
   R_f[1,15] := 0.1695628;
   R_f[2,0] := 0.8806943;
   R_f[2,1] := -0.4307577;
   R_f[2,2] := -0.285418;
   R_f[2,3] := 0.7795734;
   R_f[2,4] := 0.49964;
   R_f[2,5] := 0.1542652;
   R_f[2,6] := 0.2286351;
   R_f[2,7] := -0.7402638;
   R_f[2,8] := -0.6850481;
   R_f[2,9] := -0.3444061;
   R_f[2,10] := -0.5146202;
   R_f[2,11] := 0.5203135;
   R_f[2,12] := -0.2921089;
   R_f[2,13] := -0.7581262;
   R_f[2,14] := 0.2400508;
   R_f[2,15] := 0.06470054;
   R_f[3,0] := -1.016384;
   R_f[3,1] := -0.01572494;
   R_f[3,2] := 1.122687;
   R_f[3,3] := -1.076523;
   R_f[3,4] := -0.2219028;
   R_f[3,5] := 0.3841916;
   R_f[3,6] := 0.6512823;
   R_f[3,7] := 1.68439;
   R_f[3,8] := 0.7787917;
   R_f[3,9] := -0.1303423;
   R_f[3,10] := 0.1025792;
   R_f[3,11] := 0.0630113;
   R_f[3,12] := -0.2613996;
   R_f[3,13] := 0.08574831;
   R_f[3,14] := 0.5817915;
   R_f[3,15] := -0.1694773;
   R_f[4,0] := -0.09817147;
   R_f[4,1] := -0.8673013;
   R_f[4,2] := 0.1123603;
   R_f[4,3] := -0.05304767;
   R_f[4,4] := -0.1617602;
   R_f[4,5] := -0.4315653;
   R_f[4,6] := -0.1545042;
   R_f[4,7] := -0.04651795;
   R_f[4,8] := -0.7793221;
   R_f[4,9] := 0.2078234;
   R_f[4,10] := 0.1676973;
   R_f[4,11] := 0.3325663;
   R_f[4,12] := 0.157971;
   R_f[4,13] := 0.7362291;
   R_f[4,14] := 0.0176266;
   R_f[4,15] := -0.6734453;
   R_f[5,0] := 1.169603;
   R_f[5,1] := -0.73158;
   R_f[5,2] := 0.4122632;
   R_f[5,3] := 0.02196453;
   R_f[5,4] := 0.3548708;
   R_f[5,5] := 0.1889586;
   R_f[5,6] := 0.3045126;
   R_f[5,7] := 0.9211732;
   R_f[5,8] := -0.4857724;
   R_f[5,9] := -0.9820208;
   R_f[5,10] := -0.5130315;
   R_f[5,11] := 0.2623543;
   R_f[5,12] := -0.2203466;
   R_f[5,13] := -1.837646;
   R_f[5,14] := -0.6587409;
   R_f[5,15] := -0.2930804;
   R_f[6,0] := -0.3989139;
   R_f[6,1] := -0.7530556;
   R_f[6,2] := 1.695848;
   R_f[6,3] := -0.1637086;
   R_f[6,4] := 0.2540572;
   R_f[6,5] := 0.02853256;
   R_f[6,6] := 0.1514727;
   R_f[6,7] := -1.134142;
   R_f[6,8] := -0.9914478;
   R_f[6,9] := -0.4490964;
   R_f[6,10] := -0.6475779;
   R_f[6,11] := -0.02062916;
   R_f[6,12] := 0.3351462;
   R_f[6,13] := 0.3090186;
   R_f[6,14] := 0.6139765;
   R_f[6,15] := 0.7687923;
   R_f[7,0] := -0.2705219;
   R_f[7,1] := 0.04162847;
   R_f[7,2] := 3.147241;
   R_f[7,3] := -0.331195;
   R_f[7,4] := -0.5884408;
   R_f[7,5] := -0.3636526;
   R_f[7,6] := -0.9163497;
   R_f[7,7] := 0.3539489;
   R_f[7,8] := 0.2825061;
   R_f[7,9] := 0.493275;
   R_f[7,10] := 1.353475;
   R_f[7,11] := -1.124487;
   R_f[7,12] := -0.5918967;
   R_f[7,13] := 1.290014;
   R_f[7,14] := -0.550961;
   R_f[7,15] := 0.8665411;
   R_f[8,0] := 0.3655965;
   R_f[8,1] := -1.387398;
   R_f[8,2] := 0.6403066;
   R_f[8,3] := 0.4521842;
   R_f[8,4] := 0.426568;
   R_f[8,5] := -0.3468258;
   R_f[8,6] := -1.100012;
   R_f[8,7] := -0.6693547;
   R_f[8,8] := -3.069017;
   R_f[8,9] := 0.1657671;
   R_f[8,10] := 0.784942;
   R_f[8,11] := -0.4345917;
   R_f[8,12] := -1.434882;
   R_f[8,13] := 0.1338141;
   R_f[8,14] := -0.793483;
   R_f[8,15] := -0.2249214;
   R_f[9,0] := -0.152597;
   R_f[9,1] := -1.499914;
   R_f[9,2] := 1.108761;
   R_f[9,3] := -0.5297781;
   R_f[9,4] := -0.6886869;
   R_f[9,5] := -1.672909;
   R_f[9,6] := 2.633435;
   R_f[9,7] := -1.828544;
   R_f[9,8] := -0.740662;
   R_f[9,9] := 1.526205;
   R_f[9,10] := 0.4746018;
   R_f[9,11] := 1.381489;
   R_f[9,12] := -0.6054185;
   R_f[9,13] := 0.7926679;
   R_f[9,14] := 0.3271781;
   R_f[9,15] := -1.000112;
   R_f[10,0] := 2.164407;
   R_f[10,1] := -0.6995372;
   R_f[10,2] := 0.6653332;
   R_f[10,3] := 1.181759;
   R_f[10,4] := -0.2965346;
   R_f[10,5] := -0.1037577;
   R_f[10,6] := 0.02757812;
   R_f[10,7] := -0.9681873;
   R_f[10,8] := -0.4607585;
   R_f[10,9] := -0.5446746;
   R_f[10,10] := 0.780597;
   R_f[10,11] := -0.7688502;
   R_f[10,12] := -1.056067;
   R_f[10,13] := -0.1988855;
   R_f[10,14] := 0.01456859;
   R_f[10,15] := 0.3702135;
   R_f[11,0] := 0.2434937;
   R_f[11,1] := -0.1798942;
   R_f[11,2] := 0.2355876;
   R_f[11,3] := -0.6682997;
   R_f[11,4] := -0.5007147;
   R_f[11,5] := -0.5791205;
   R_f[11,6] := 0.1253008;
   R_f[11,7] := -0.7620748;
   R_f[11,8] := -0.5787513;
   R_f[11,9] := 0.0264844;
   R_f[11,10] := 0.4317927;
   R_f[11,11] := -1.222577;
   R_f[11,12] := -0.03755289;
   R_f[11,13] := -0.1228497;
   R_f[11,14] := 0.0646783;
   R_f[11,15] := 0.2649987;
   R_f[12,0] := -0.02412502;
   R_f[12,1] := -0.4178893;
   R_f[12,2] := 0.2250565;
   R_f[12,3] := 0.2468531;
   R_f[12,4] := -0.2603359;
   R_f[12,5] := 0.5588626;
   R_f[12,6] := 0.3501927;
   R_f[12,7] := 0.0646469;
   R_f[12,8] := 0.3895332;
   R_f[12,9] := 0.409056;
   R_f[12,10] := 0.161415;
   R_f[12,11] := -0.05112006;
   R_f[12,12] := 1.493768;
   R_f[12,13] := 0.3131461;
   R_f[12,14] := 0.4573432;
   R_f[12,15] := 0.3800302;
   R_f[13,0] := 0.5914586;
   R_f[13,1] := -0.351166;
   R_f[13,2] := 0.8291268;
   R_f[13,3] := 0.2013447;
   R_f[13,4] := 0.82876;
   R_f[13,5] := 0.8977232;
   R_f[13,6] := 1.657781;
   R_f[13,7] := 0.4952854;
   R_f[13,8] := -0.8510268;
   R_f[13,9] := -0.7816306;
   R_f[13,10] := 0.3712052;
   R_f[13,11] := 0.7794952;
   R_f[13,12] := -0.1510022;
   R_f[13,13] := -0.1749281;
   R_f[13,14] := -0.00674355;
   R_f[13,15] := -0.6594451;
   R_f[14,0] := -0.03948923;
   R_f[14,1] := -0.3682528;
   R_f[14,2] := 1.244398;
   R_f[14,3] := -0.5374001;
   R_f[14,4] := -0.4286888;
   R_f[14,5] := 0.2608948;
   R_f[14,6] := 0.4886785;
   R_f[14,7] := 1.195282;
   R_f[14,8] := 0.1545673;
   R_f[14,9] := -1.140402;
   R_f[14,10] := 0.05182516;
   R_f[14,11] := -0.2172662;
   R_f[14,12] := 0.1702152;
   R_f[14,13] := -0.6474801;
   R_f[14,14] := 1.387721;
   R_f[14,15] := 0.2322865;
   R_f[15,0] := 0.3153065;
   R_f[15,1] := -0.9808237;
   R_f[15,2] := 0.2264991;
   R_f[15,3] := -0.2976737;
   R_f[15,4] := 0.5468484;
   R_f[15,5] := 0.7780918;
   R_f[15,6] := 2.003952;
   R_f[15,7] := 2.355743;
   R_f[15,8] := -0.1702361;
   R_f[15,9] := -0.381211;
   R_f[15,10] := 1.069254;
   R_f[15,11] := -0.3054578;
   R_f[15,12] := -0.4347287;
   R_f[15,13] := -1.114827;
   R_f[15,14] := 0.3245434;
   R_f[15,15] := -1.337709;
   R_g[0,0] := -2.805433;
   R_g[0,1] := 0.09675837;
   R_g[0,2] := 0.04763355;
   R_g[0,3] := 0.1613498;
   R_g[0,4] := -0.04916951;
   R_g[0,5] := 0.06786807;
   R_g[0,6] := 0.07195669;
   R_g[0,7] := 0.1879627;
   R_g[0,8] := 0.02096096;
   R_g[0,9] := -0.05091592;
   R_g[0,10] := 0.1711352;
   R_g[0,11] := 0.09710391;
   R_g[0,12] := -0.1928508;
   R_g[0,13] := 0.04608029;
   R_g[0,14] := 0.3775772;
   R_g[0,15] := -0.05004899;
   R_g[1,0] := 0.08712953;
   R_g[1,1] := -1.281738;
   R_g[1,2] := 0.486291;
   R_g[1,3] := -0.1018547;
   R_g[1,4] := 0.5911466;
   R_g[1,5] := 0.3826247;
   R_g[1,6] := 0.04029783;
   R_g[1,7] := 0.06582787;
   R_g[1,8] := -0.06752597;
   R_g[1,9] := -0.2294858;
   R_g[1,10] := -0.1253151;
   R_g[1,11] := -0.2067355;
   R_g[1,12] := -0.05208173;
   R_g[1,13] := 0.1810765;
   R_g[1,14] := 0.05905702;
   R_g[1,15] := -0.06634986;
   R_g[2,0] := -0.2549139;
   R_g[2,1] := -0.05303259;
   R_g[2,2] := -3.258265;
   R_g[2,3] := 0.2239036;
   R_g[2,4] := 0.08010214;
   R_g[2,5] := 0.1251935;
   R_g[2,6] := -0.1281362;
   R_g[2,7] := 0.03709217;
   R_g[2,8] := -0.0533942;
   R_g[2,9] := -0.1838315;
   R_g[2,10] := 0.01583981;
   R_g[2,11] := 0.1206139;
   R_g[2,12] := 0.02361463;
   R_g[2,13] := 0.1162473;
   R_g[2,14] := 0.1685608;
   R_g[2,15] := -0.04670952;
   R_g[3,0] := -0.3499806;
   R_g[3,1] := 0.7145555;
   R_g[3,2] := -0.7979932;
   R_g[3,3] := -2.84151;
   R_g[3,4] := 0.1580465;
   R_g[3,5] := -0.08033045;
   R_g[3,6] := -0.1452473;
   R_g[3,7] := 0.2225952;
   R_g[3,8] := 0.07427457;
   R_g[3,9] := 0.3725025;
   R_g[3,10] := -0.308892;
   R_g[3,11] := -0.2322429;
   R_g[3,12] := 0.6733903;
   R_g[3,13] := 0.1802014;
   R_g[3,14] := -0.04057474;
   R_g[3,15] := -0.1780594;
   R_g[4,0] := 0.4558564;
   R_g[4,1] := 0.2691017;
   R_g[4,2] := 0.2479934;
   R_g[4,3] := 0.1830495;
   R_g[4,4] := -2.643592;
   R_g[4,5] := -0.1854873;
   R_g[4,6] := 0.5796254;
   R_g[4,7] := -0.2360368;
   R_g[4,8] := 0.3996172;
   R_g[4,9] := -0.08552616;
   R_g[4,10] := -0.3547961;
   R_g[4,11] := 0.02176627;
   R_g[4,12] := -0.1695444;
   R_g[4,13] := -0.6054811;
   R_g[4,14] := 0.05480947;
   R_g[4,15] := 0.2614591;
   R_g[5,0] := 0.09851117;
   R_g[5,1] := 0.05978253;
   R_g[5,2] := -0.2238024;
   R_g[5,3] := 0.06287329;
   R_g[5,4] := 0.2952785;
   R_g[5,5] := -6.417284;
   R_g[5,6] := -0.01966351;
   R_g[5,7] := 0.08289347;
   R_g[5,8] := 0.2335418;
   R_g[5,9] := 0.4640638;
   R_g[5,10] := -0.5190796;
   R_g[5,11] := -0.3999299;
   R_g[5,12] := 0.3029557;
   R_g[5,13] := 0.06150499;
   R_g[5,14] := -1.054952;
   R_g[5,15] := -0.08431676;
   R_g[6,0] := -0.1025641;
   R_g[6,1] := 0.05051776;
   R_g[6,2] := 0.0306027;
   R_g[6,3] := 0.06608646;
   R_g[6,4] := -0.05028161;
   R_g[6,5] := -0.1038706;
   R_g[6,6] := -3.13754;
   R_g[6,7] := -0.1565541;
   R_g[6,8] := 0.03909466;
   R_g[6,9] := -0.03506904;
   R_g[6,10] := 0.0048442;
   R_g[6,11] := -0.1906409;
   R_g[6,12] := 0.330723;
   R_g[6,13] := -0.06755624;
   R_g[6,14] := -0.1569814;
   R_g[6,15] := -0.3220711;
   R_g[7,0] := 0.07863971;
   R_g[7,1] := -0.1875482;
   R_g[7,2] := -0.2537812;
   R_g[7,3] := -0.08824939;
   R_g[7,4] := -0.1294116;
   R_g[7,5] := 0.2885412;
   R_g[7,6] := 0.1121606;
   R_g[7,7] := -3.136752;
   R_g[7,8] := -0.08472223;
   R_g[7,9] := 0.00790842;
   R_g[7,10] := -0.1138648;
   R_g[7,11] := -0.05684523;
   R_g[7,12] := 0.1106585;
   R_g[7,13] := -0.07569506;
   R_g[7,14] := 0.4233017;
   R_g[7,15] := -0.1342552;
   R_g[8,0] := 0.08961181;
   R_g[8,1] := 0.4651947;
   R_g[8,2] := -0.3656231;
   R_g[8,3] := 0.2111352;
   R_g[8,4] := -0.00757714;
   R_g[8,5] := -0.2639286;
   R_g[8,6] := 0.1638752;
   R_g[8,7] := -0.4058702;
   R_g[8,8] := -2.934379;
   R_g[8,9] := 0.08376594;
   R_g[8,10] := -0.2960652;
   R_g[8,11] := 0.01828978;
   R_g[8,12] := 0.2524873;
   R_g[8,13] := -0.3134462;
   R_g[8,14] := -0.01567479;
   R_g[8,15] := 0.05443858;
   R_g[9,0] := -0.1509652;
   R_g[9,1] := -0.2985869;
   R_g[9,2] := 0.1976654;
   R_g[9,3] := -0.1125526;
   R_g[9,4] := -0.1207261;
   R_g[9,5] := 0.337102;
   R_g[9,6] := 0.2015858;
   R_g[9,7] := -0.1138979;
   R_g[9,8] := -0.08645659;
   R_g[9,9] := -4.490891;
   R_g[9,10] := 0.03153508;
   R_g[9,11] := 0.1759175;
   R_g[9,12] := -0.00816477;
   R_g[9,13] := -0.09244221;
   R_g[9,14] := -0.1702342;
   R_g[9,15] := 0.4290646;
   R_g[10,0] := -0.3885716;
   R_g[10,1] := 0.0643687;
   R_g[10,2] := -0.1564249;
   R_g[10,3] := -0.1040558;
   R_g[10,4] := 0.1323418;
   R_g[10,5] := 0.1366159;
   R_g[10,6] := 0.04957649;
   R_g[10,7] := 0.0648922;
   R_g[10,8] := 0.1469345;
   R_g[10,9] := -0.01300282;
   R_g[10,10] := -1.928301;
   R_g[10,11] := 0.3004588;
   R_g[10,12] := 0.2731377;
   R_g[10,13] := 0.02955168;
   R_g[10,14] := -0.07842075;
   R_g[10,15] := 0.05753986;
   R_g[11,0] := -0.2097152;
   R_g[11,1] := 0.7307096;
   R_g[11,2] := -0.503158;
   R_g[11,3] := 0.205001;
   R_g[11,4] := -0.01089373;
   R_g[11,5] := 0.16405;
   R_g[11,6] := 0.1890694;
   R_g[11,7] := 0.03491729;
   R_g[11,8] := -0.01610962;
   R_g[11,9] := 0.2807466;
   R_g[11,10] := 0.02013272;
   R_g[11,11] := -4.203784;
   R_g[11,12] := 0.2934183;
   R_g[11,13] := 0.1436955;
   R_g[11,14] := -0.41985;
   R_g[11,15] := 0.0576296;
   R_g[12,0] := -0.03705381;
   R_g[12,1] := -0.3112487;
   R_g[12,2] := 0.6347389;
   R_g[12,3] := 0.08633271;
   R_g[12,4] := -0.1792604;
   R_g[12,5] := 0.317774;
   R_g[12,6] := -0.1986456;
   R_g[12,7] := -0.1977208;
   R_g[12,8] := 0.1422061;
   R_g[12,9] := -0.2642545;
   R_g[12,10] := 0.07095157;
   R_g[12,11] := 0.5123266;
   R_g[12,12] := -3.63069;
   R_g[12,13] := -0.1175799;
   R_g[12,14] := 0.2990645;
   R_g[12,15] := -0.02980175;
   R_g[13,0] := 0.00863379;
   R_g[13,1] := 0.03295338;
   R_g[13,2] := -0.3002235;
   R_g[13,3] := 0.1032756;
   R_g[13,4] := -0.1160595;
   R_g[13,5] := 0.031227;
   R_g[13,6] := 0.6257741;
   R_g[13,7] := 0.4343066;
   R_g[13,8] := 0.1252338;
   R_g[13,9] := 0.1524162;
   R_g[13,10] := -0.2399488;
   R_g[13,11] := -0.0243434;
   R_g[13,12] := 0.07577311;
   R_g[13,13] := -2.642776;
   R_g[13,14] := -0.7371749;
   R_g[13,15] := -0.08735505;
   R_g[14,0] := -0.171414;
   R_g[14,1] := 0.2261713;
   R_g[14,2] := -0.3317359;
   R_g[14,3] := 0.0877693;
   R_g[14,4] := 0.1621639;
   R_g[14,5] := 0.2182705;
   R_g[14,6] := 0.04451356;
   R_g[14,7] := 0.03265934;
   R_g[14,8] := -0.136193;
   R_g[14,9] := 0.1847814;
   R_g[14,10] := -0.0108934;
   R_g[14,11] := -0.2341314;
   R_g[14,12] := 0.1122679;
   R_g[14,13] := 0.2223738;
   R_g[14,14] := -2.0286;
   R_g[14,15] := -0.01800863;
   R_g[15,0] := 0.3883483;
   R_g[15,1] := -0.1211964;
   R_g[15,2] := -0.4713392;
   R_g[15,3] := 0.02589257;
   R_g[15,4] := -0.1296599;
   R_g[15,5] := -0.2871422;
   R_g[15,6] := 0.6408823;
   R_g[15,7] := 0.4650818;
   R_g[15,8] := -0.1301513;
   R_g[15,9] := 0.1214571;
   R_g[15,10] := 0.3844216;
   R_g[15,11] := -0.5117303;
   R_g[15,12] := -0.03178278;
   R_g[15,13] := -0.2080431;
   R_g[15,14] := 0.6247337;
   R_g[15,15] := -3.379229;
   R_o[0,0] := -0.148473;
   R_o[0,1] := -0.7470531;
   R_o[0,2] := 0.337931;
   R_o[0,3] := 0.4881276;
   R_o[0,4] := -0.5424621;
   R_o[0,5] := 0.2365883;
   R_o[0,6] := 0.3687733;
   R_o[0,7] := -0.04479291;
   R_o[0,8] := 0.04525228;
   R_o[0,9] := -0.06947453;
   R_o[0,10] := -0.2940823;
   R_o[0,11] := -0.6614071;
   R_o[0,12] := -0.09016941;
   R_o[0,13] := -0.2445324;
   R_o[0,14] := 0.4173301;
   R_o[0,15] := 0.1152808;
   R_o[1,0] := -0.2253625;
   R_o[1,1] := -2.687598;
   R_o[1,2] := 0.7825195;
   R_o[1,3] := 0.3311445;
   R_o[1,4] := -0.6487191;
   R_o[1,5] := -0.1774464;
   R_o[1,6] := -0.6072173;
   R_o[1,7] := -0.9984445;
   R_o[1,8] := 0.693763;
   R_o[1,9] := -0.04945409;
   R_o[1,10] := 0.1380522;
   R_o[1,11] := 0.2601311;
   R_o[1,12] := -0.5988305;
   R_o[1,13] := -1.649512;
   R_o[1,14] := -0.06540374;
   R_o[1,15] := -0.683998;
   R_o[2,0] := 0.1426505;
   R_o[2,1] := -0.7636122;
   R_o[2,2] := 0.6522185;
   R_o[2,3] := -0.01308598;
   R_o[2,4] := -0.3956572;
   R_o[2,5] := -0.1286385;
   R_o[2,6] := 0.1117783;
   R_o[2,7] := -0.1965184;
   R_o[2,8] := 0.445568;
   R_o[2,9] := -0.3197942;
   R_o[2,10] := 0.1024574;
   R_o[2,11] := -0.3961471;
   R_o[2,12] := -0.1107483;
   R_o[2,13] := -0.7957024;
   R_o[2,14] := 0.2206428;
   R_o[2,15] := 0.2849079;
   R_o[3,0] := 0.103478;
   R_o[3,1] := -0.3351506;
   R_o[3,2] := 0.1007192;
   R_o[3,3] := 0.2476437;
   R_o[3,4] := -0.3063624;
   R_o[3,5] := -0.02347863;
   R_o[3,6] := 0.6147529;
   R_o[3,7] := 0.05460903;
   R_o[3,8] := -0.09153262;
   R_o[3,9] := -0.07667586;
   R_o[3,10] := 0.1709715;
   R_o[3,11] := -0.847174;
   R_o[3,12] := 0.01488861;
   R_o[3,13] := 0.01246201;
   R_o[3,14] := 0.785248;
   R_o[3,15] := -0.2429155;
   R_o[4,0] := 0.7403428;
   R_o[4,1] := -1.202408;
   R_o[4,2] := -0.01728833;
   R_o[4,3] := -0.2675001;
   R_o[4,4] := 0.4232838;
   R_o[4,5] := -0.1884229;
   R_o[4,6] := -0.4024306;
   R_o[4,7] := 0.6314479;
   R_o[4,8] := -1.543486;
   R_o[4,9] := 0.5625891;
   R_o[4,10] := -0.4602357;
   R_o[4,11] := -0.7463102;
   R_o[4,12] := 0.01794407;
   R_o[4,13] := 0.6175683;
   R_o[4,14] := -0.4240062;
   R_o[4,15] := -0.3216551;
   R_o[5,0] := -1.608714;
   R_o[5,1] := -0.8543944;
   R_o[5,2] := 0.1236723;
   R_o[5,3] := 0.3216394;
   R_o[5,4] := -0.4782757;
   R_o[5,5] := 3.932515;
   R_o[5,6] := -0.1368901;
   R_o[5,7] := 1.26777;
   R_o[5,8] := -0.6972287;
   R_o[5,9] := -0.6138417;
   R_o[5,10] := 0.9199839;
   R_o[5,11] := -0.644981;
   R_o[5,12] := -0.2947383;
   R_o[5,13] := -1.30751;
   R_o[5,14] := 0.8453699;
   R_o[5,15] := 1.6406;
   R_o[6,0] := 0.02413699;
   R_o[6,1] := -0.7911229;
   R_o[6,2] := -0.1035878;
   R_o[6,3] := -0.345346;
   R_o[6,4] := 0.4822478;
   R_o[6,5] := -0.5942275;
   R_o[6,6] := 0.5900132;
   R_o[6,7] := 0.05578557;
   R_o[6,8] := -0.1626476;
   R_o[6,9] := -0.5127108;
   R_o[6,10] := 0.395417;
   R_o[6,11] := -0.5891114;
   R_o[6,12] := -0.04537732;
   R_o[6,13] := 0.2378311;
   R_o[6,14] := 0.5396131;
   R_o[6,15] := 0.6403692;
   R_o[7,0] := 0.1401259;
   R_o[7,1] := -1.107673;
   R_o[7,2] := 0.449949;
   R_o[7,3] := 0.1980791;
   R_o[7,4] := -0.1763375;
   R_o[7,5] := -0.02624386;
   R_o[7,6] := 0.6654956;
   R_o[7,7] := 0.8419639;
   R_o[7,8] := 0.07700922;
   R_o[7,9] := 0.585766;
   R_o[7,10] := 0.117281;
   R_o[7,11] := -0.205901;
   R_o[7,12] := -0.1026604;
   R_o[7,13] := 0.1098014;
   R_o[7,14] := 0.8365094;
   R_o[7,15] := 0.4066797;
   R_o[8,0] := 0.1040777;
   R_o[8,1] := -1.388284;
   R_o[8,2] := 0.5748492;
   R_o[8,3] := -0.3209612;
   R_o[8,4] := -1.21653;
   R_o[8,5] := -0.1644516;
   R_o[8,6] := 0.521858;
   R_o[8,7] := 2.041153;
   R_o[8,8] := -2.922855;
   R_o[8,9] := -0.6003711;
   R_o[8,10] := -0.1361148;
   R_o[8,11] := -0.102449;
   R_o[8,12] := -0.5256941;
   R_o[8,13] := -0.3414919;
   R_o[8,14] := 0.9229004;
   R_o[8,15] := -0.1494768;
   R_o[9,0] := 0.9020318;
   R_o[9,1] := -1.182273;
   R_o[9,2] := 0.7037838;
   R_o[9,3] := -0.07063206;
   R_o[9,4] := -0.4500138;
   R_o[9,5] := 0.3359483;
   R_o[9,6] := 0.9089686;
   R_o[9,7] := -0.1131394;
   R_o[9,8] := 0.06154737;
   R_o[9,9] := -3.070117;
   R_o[9,10] := 0.2449786;
   R_o[9,11] := -0.03553757;
   R_o[9,12] := -0.3328317;
   R_o[9,13] := 0.3393808;
   R_o[9,14] := 0.4877961;
   R_o[9,15] := 0.9906611;
   R_o[10,0] := 0.3674809;
   R_o[10,1] := -0.4065204;
   R_o[10,2] := 0.3212383;
   R_o[10,3] := 0.1469396;
   R_o[10,4] := -0.8636696;
   R_o[10,5] := 0.4387633;
   R_o[10,6] := -0.3679813;
   R_o[10,7] := -0.3709672;
   R_o[10,8] := 0.8587736;
   R_o[10,9] := -0.4086122;
   R_o[10,10] := 1.240259;
   R_o[10,11] := -0.5606848;
   R_o[10,12] := -0.1593753;
   R_o[10,13] := -0.5910825;
   R_o[10,14] := 0.8222155;
   R_o[10,15] := 0.07025416;
   R_o[11,0] := -0.283336;
   R_o[11,1] := -0.8366182;
   R_o[11,2] := 0.2441355;
   R_o[11,3] := 0.1767131;
   R_o[11,4] := -0.4013823;
   R_o[11,5] := 0.1624961;
   R_o[11,6] := 0.590718;
   R_o[11,7] := 1.182436;
   R_o[11,8] := -0.1144639;
   R_o[11,9] := -0.459346;
   R_o[11,10] := 0.4479548;
   R_o[11,11] := 1.724371;
   R_o[11,12] := -0.6445624;
   R_o[11,13] := -0.2646877;
   R_o[11,14] := 1.049319;
   R_o[11,15] := 1.146086;
   R_o[12,0] := 0.06811738;
   R_o[12,1] := -0.8294082;
   R_o[12,2] := 0.04298686;
   R_o[12,3] := 0.1884655;
   R_o[12,4] := -0.4888053;
   R_o[12,5] := 0.06246455;
   R_o[12,6] := 0.5130124;
   R_o[12,7] := 0.01585177;
   R_o[12,8] := -0.3286436;
   R_o[12,9] := -0.1914053;
   R_o[12,10] := 0.3550029;
   R_o[12,11] := -0.6732444;
   R_o[12,12] := -0.1367572;
   R_o[12,13] := 0.1686232;
   R_o[12,14] := 0.7652449;
   R_o[12,15] := 0.1804299;
   R_o[13,0] := 1.529198;
   R_o[13,1] := -2.016652;
   R_o[13,2] := 0.07069629;
   R_o[13,3] := 0.5932482;
   R_o[13,4] := -0.01248456;
   R_o[13,5] := 0.1003619;
   R_o[13,6] := 0.9069089;
   R_o[13,7] := 0.4181206;
   R_o[13,8] := -0.1110177;
   R_o[13,9] := -0.4146234;
   R_o[13,10] := 0.3274502;
   R_o[13,11] := 0.09499595;
